(* IEC 61131-3 sources: 2026_Projet_YGO_ExcavatriceDragage/CODE/M_MAIN (part 2) *)

M1WinchSensors.CablePosM          := PRG_02_Acquisition.Data.EncoderM1.Measurement.CablePosM;
M1WinchSensors.Homed              := PRG_02_Acquisition.Data.EncoderM1.Homed;
M1WinchSensors.HomingSuspect      := PRG_02_Acquisition.Data.EncoderM1.HomingSuspect;
M1WinchSensors.ContactorsAllOff   := PRG_02_Acquisition.HwIn.Winch.M1_ContactorsReleased_DI;
M1WinchSensors.MeasuredSpeedBand  := instWinchLoadEstimatorM1.SpeedBand;
// Garde-fou vitesse mesuree : DESACTIVE par defaut (AF_Partie-10 §9bis, FB_Winch_v2.1 /
// FB_SpeedStep_v1.0 SpeedGuardEnable := FALSE). Le TRUE code en dur etait un reste de
// mise en service : il rendait la capacite de palier otage de instWinchSync (tout ecart
// sync -> SpeedGuardReady=FALSE -> clamp palier 1, y compris en montee).
// ⚠️ DETTE SAFETY -S5 : le garde-fou vitesse mesuree est HORS SERVICE. Le FB de
// gouvernance nominale annonce (FB_WinchRateInterlock) n'existe PAS dans CODE/.
// Decision : risque ACTE et documente — la surveillance survitesse reelle est portee par
// FB_Safety_Winch (gelee : harnais VAR_IN_OUT indisponible). Ne PAS armer une
// survitesse sur une table non prouvee. A re-trancher a la livraison .
// ⚠️ tache est BLOQUE (contrat C4 TASK_CONTRACT_AUTORITE_2_INTERLOCKS.yaml,
// ARRET VALIDATION HUMAINE requis : autorite, T_max/DropConfirmDelay, classification
// Fault.Error, argument PLr ; prerequis// non livres). Ne PAS creer
// FB_WinchRateInterlock hors de ce contrat — la logique de garde-fou existe deja dans
// FB_Winch §5 et reste volontairement desactivee (SpeedGuardEnable := FALSE) tant que la
// table SpeedBandMaxMps n'est pas validee en charge reelle (AF-10 §7.3 TBD).
M1WinchSensors.SpeedGuardEnable   := FALSE;
M1WinchSensors.SpeedGuardReady    := NOT instWinchSync.Fault.Error;

M1WinchCfg.SpeedStepTable         := _WinchSpeedStepTable;
M1WinchCfg.SlowdownDistanceTop_M  := _CommunCfgPersist.WinchSlowdownDistanceTop_M;
M1WinchCfg.SlowdownDistanceBottom_M := _CommunCfgPersist.WinchSlowdownDistanceBottom_M;
M1WinchCfg.SlowdownMaxStep        := _CommunCfgPersist.WinchSlowdownMaxStep;
// Cadence/interlocks : descente normale 500 ms, inversion vers descente 500 ms,
// montee normale 700 ms, inversion vers montee 800 ms.
// Champs non portes par la persistante -> assignes explicitement (le defaut de type n'est
// pas applique au runtime pour ce VAR local de struct). 0,7 s montee / 0,5 s descente.
M1WinchCfg.DirectionInterlockDelayAscent  := T#800ms;
M1WinchCfg.DirectionInterlockDelayDescent := T#500ms;
M1WinchCfg.StepRampDelayAscent    := T#700ms;
M1WinchCfg.StepRampDelayDescent   := T#500ms;

instWinchM1(
    Enable                  := (PRG_03_Modes_Cycle.Data.Auth.Mode <> E_Mode.DISABLE) AND NOT PRG_03_Modes_Cycle.Data.Auth.InhibitM1,
    Reset                   := PRG_07_Supervision.FaultMachineReset_IHM,
    PowerContactorEngaged   := PRG_02_Acquisition.HwIn.Machine.PowerContactorEngaged_DI,
    SafeStop                := SafeStopM1_Active,
    DescendPermit           := EffectivePermitM1_Descend,
    AscentPermit            := EffectivePermitM1_Ascent,
    WinchRequest            := ReqM1Winch,
    Sensors                 := M1WinchSensors,
    Config                  := M1WinchCfg,
    // ContactorFeedback (n°3 de la matrice) et Global — sans gate de mode (dérogation MES 2026).
    BypassContactorCheck    := (GVL_IHM.M1TreuilRetenue.Bypass.Global OR GVL_IHM.M1TreuilRetenue.Bypass.ContactorFeedback),
    BypassGlobal            := GVL_IHM.M1TreuilRetenue.Bypass.Global
);

// --- M2 : assemblage des structs ---
ReqM2Winch.RunRequest               := M2LogicRunRequest;
ReqM2Winch.ReqAscent                := M2LogicReqAscent;
ReqM2Winch.ReqDescend               := M2LogicReqDescend;
ReqM2Winch.SpeedStepReq             := M2LogicRequestStepTgt;
// Clamp de palier agrégé en §5ter : bornes communes M1=M2 (CommonMaxStep*) puis
// M2-propre (M2MaxStep*) — M2_BucketJogLimit / ManualBucketLimitsActive ne réduisent
// jamais M1 (pilotage unitaire M2). BucketNotClosedAscentCapStep1 /
// SlackCableAscentCapStep1 : réduisent M1 aussi UNIQUEMENT en pilotage couplé
// (CoupledBoth) — les 2 treuils liés doivent rester au même palier.
// D13 : reconstruction de table M2 supprimée — le clamp M2MaxStep* := 1 suffit
// (StepNumber ≤ 1 → seuls les états P1 sont commandés).
ReqM2Winch.MaxStepUp                := M2MaxStepUp;
ReqM2Winch.MaxStepDown              := M2MaxStepDown;
// Plancher palier descente plongée Kobold : plancher M2-propre agrégé en §5ter, injecté
// sur la cible (jamais sur StepNumber). Aucun effet si StartStop=FALSE.
ReqM2Winch.MinStepDown              := M2MinStepDown;
ReqM2Winch.HomingApproachActive     := PRG_03_Modes_Cycle.Data.Auth.HomingApproachEnable;
// Même limite haute active que FB_Safety_Winch (M2_LimitShift conservé).
ReqM2Winch.TopLimitM                := TopLimitM2_M;
ReqM2Winch.BottomLimitM             := BottomLimitM2_Active;
ReqM2Winch.SyncCoupled              := instWinchSync.SyncActive;

// === ATOMICITE DU DEMARRAGE COUPLE (volet M2, symetrique du volet M1 ~ligne 1225) ===
// Meme verrou : en intention both, si l'un des deux treuils n'est pas pret, on fige AUSSI
// la commande finale M2. Cas symetrique du REX : M2 relance seul pendant que M1 est en
// dead-time D18 -> cable qui file. On fige M2 UNIQUEMENT si M1 est le treuil pas pret.
IF NOT MaintN2 AND WinchBothMotionActive AND (instWinchM1.DirectionChangePending OR instWinchM1.Fault.Latched) THEN
    ReqM2Winch.RunRequest := FALSE; ReqM2Winch.ReqAscent := FALSE; ReqM2Winch.ReqDescend := FALSE; ReqM2Winch.SpeedStepReq := 0;
END_IF;

M2WinchSensors.CablePosM          := PRG_02_Acquisition.Data.EncoderM2.Measurement.CablePosM;
M2WinchSensors.Homed              := PRG_02_Acquisition.Data.EncoderM2.Homed;
M2WinchSensors.HomingSuspect      := PRG_02_Acquisition.Data.EncoderM2.HomingSuspect;
M2WinchSensors.ContactorsAllOff   := PRG_02_Acquisition.HwIn.Winch.M2_ContactorsReleased_DI;
M2WinchSensors.MeasuredSpeedBand  := instWinchLoadEstimatorM2.SpeedBand;
// Garde-fou vitesse mesuree : DESACTIVE par defaut (idem M1 ci-dessus, AF_Partie-10 §9bis).
M2WinchSensors.SpeedGuardEnable   := FALSE;
M2WinchSensors.SpeedGuardReady    := NOT instWinchSync.Fault.Error;

M2WinchCfg.SpeedStepTable         := _WinchSpeedStepTable;
M2WinchCfg.SlowdownDistanceTop_M  := _CommunCfgPersist.WinchSlowdownDistanceTop_M;
M2WinchCfg.SlowdownDistanceBottom_M := _CommunCfgPersist.WinchSlowdownDistanceBottom_M;
M2WinchCfg.SlowdownMaxStep        := _CommunCfgPersist.WinchSlowdownMaxStep;
// Cadence/interlocks identiques M1 : descente normale 500 ms, inversion vers descente
// 500 ms, montee normale 700 ms, inversion vers montee 800 ms.
M2WinchCfg.DirectionInterlockDelayAscent  := T#800ms;
M2WinchCfg.DirectionInterlockDelayDescent := T#500ms;
M2WinchCfg.StepRampDelayAscent    := T#700ms;
M2WinchCfg.StepRampDelayDescent   := T#500ms;

instWinchM2(
    Enable                  := (PRG_03_Modes_Cycle.Data.Auth.Mode <> E_Mode.DISABLE) AND NOT PRG_03_Modes_Cycle.Data.Auth.InhibitM2,
    Reset                   := PRG_07_Supervision.FaultMachineReset_IHM,
    PowerContactorEngaged   := PRG_02_Acquisition.HwIn.Machine.PowerContactorEngaged_DI,
    SafeStop                := SafeStopM2_Active,
    DescendPermit           := M2DescendPermitApplied,
    AscentPermit            := M2AscentPermitApplied,
    WinchRequest            := ReqM2Winch,
    Sensors                 := M2WinchSensors,
    Config                  := M2WinchCfg,
    // Idem M1 ci-dessus
    BypassContactorCheck    := (GVL_IHM.M2TreuilBenne.Bypass.Global OR GVL_IHM.M2TreuilBenne.Bypass.ContactorFeedback),
    BypassGlobal            := GVL_IHM.M2TreuilBenne.Bypass.Global
);

// Atomicite de sortie couplee : les deux FB_Winch ont maintenant traite la demande du
// scan. Leur readiness directionnelle courante est donc connue avant publication vers
// PRG_06. La barriere finale ne recevra aucun relais/contacteur tant qu'un axe attend.
WinchBothMotionReady := NOT (instWinchM1.DirectionChangePending OR instWinchM2.DirectionChangePending)
                        AND NOT instWinchM1.Fault.Latched AND NOT instWinchM2.Fault.Latched;

// ── Collecteurs passifs d'apprentissage vitesse par palier ──
// Appelés APRÈS instWinchM1/M2 : StepNumber lu = palier courant du scan (pas de lag).
// Dérivations des entrées de collecte :
//   • LoadPresent : charge présente si l'estimateur de charge (même source vitesse) estime
//     une charge >= 50 % (seuil de mise en service, à confirmer sur site).
//   • StableForLearn : treuil commandé (palier > 0) et sans défaut — conditions stables.
// Collecteur STRICTEMENT PASSIF : aucune commande moteur, aucune surveillance survitesse
// (la survitesse reste, gelée — voir bandeau §6 M1/M2 SpeedGuardEnable).
LoadPresentM1 := (instWinchLoadEstimatorM1.EstimatedLoadPct >= 50.0);
LoadPresentM2 := (instWinchLoadEstimatorM2.EstimatedLoadPct >= 50.0);
StableForLearnM1 := (instWinchM1.StepNumber > 0) AND NOT instWinchM1.Fault.Error;
StableForLearnM2 := (instWinchM2.StepNumber > 0) AND NOT instWinchM2.Fault.Error;

instWinchSpeedLearningM1(
    Enable              := (PRG_03_Modes_Cycle.Data.Auth.Mode <> E_Mode.DISABLE) AND NOT PRG_03_Modes_Cycle.Data.Auth.InhibitM1,
    LearnStart          := GVL_IHM.M1TreuilRetenue.Cmd.BtnLearnSpeed,
    WinchId             := 1,
    ReqAscent          := M1LogicReqAscent,
    ReqDescend         := M1LogicReqDescend,
    StepNumber          := instWinchM1.StepNumber,
    MeasuredSpeedMps    := PRG_02_Acquisition.Data.EncoderM1.Measurement.Speed_Mps,
    MeasuredSpeedValid  := PRG_02_Acquisition.Data.EncoderM1.Measurement.SpeedValid,
    LoadPresent         := LoadPresentM1,
    StableForLearn      := StableForLearnM1,
    Config              := _WinchSpeedLearnCfg,
    Table               := _WinchSpeedLearnTable
);

instWinchSpeedLearningM2(
    Enable              := (PRG_03_Modes_Cycle.Data.Auth.Mode <> E_Mode.DISABLE) AND NOT PRG_03_Modes_Cycle.Data.Auth.InhibitM2,
    LearnStart          := GVL_IHM.M2TreuilBenne.Cmd.BtnLearnSpeed,
    WinchId             := 2,
    ReqAscent          := M2LogicReqAscent,
    ReqDescend         := M2LogicReqDescend,
    StepNumber          := instWinchM2.StepNumber,
    MeasuredSpeedMps    := PRG_02_Acquisition.Data.EncoderM2.Measurement.Speed_Mps,
    MeasuredSpeedValid  := PRG_02_Acquisition.Data.EncoderM2.Measurement.SpeedValid,
    LoadPresent         := LoadPresentM2,
    StableForLearn      := StableForLearnM2,
    Config              := _WinchSpeedLearnCfg,
    Table               := _WinchSpeedLearnTable
);

{endregion}

{region "📤 §7 Publication demandes"}
// === 📤 §7 PUBLICATION DEMANDES BRUTES (WinchM1/M2FinalInterlockRequest) ===

WinchM1FinalInterlockRequest.Enable := TRUE;
WinchM1FinalInterlockRequest.Reset := PRG_07_Supervision.FaultMachineReset_IHM;
WinchM1FinalInterlockRequest.PowerContactorEngaged := PRG_02_Acquisition.HwIn.Machine.PowerContactorEngaged_DI;
WinchM1FinalInterlockRequest.SafeStop := SafeStopM1_Active;
// Plus de BrakeReleaseRequest/
// BrakeCommandOpenConfirmed calcules par FB_Winch — la barriere finale
// (FB_WinchOutputInterlock) recoit le retour PHYSIQUE brut directement,
// et calcule elle-meme BrakeCmd := RelayFwd OR RelayRev (voir bandeau de ce FB).
WinchM1FinalInterlockRequest.BrakeFeedback := SEL(MaintN2 OR GVL_IHM.M1TreuilRetenue.Bypass.ContactorFeedback OR GVL_IHM.M1TreuilRetenue.Bypass.Global,
                                                   PRG_02_Acquisition.HwIn.Winch.M1_BrakeIsOpen_DI,
                                                   instWinchM1.RelayFwd OR instWinchM1.RelayRev);
WinchM1FinalInterlockRequest.FwdRevSpeedFeedbackOff := SEL(MaintN2 OR GVL_IHM.M1TreuilRetenue.Bypass.ContactorFeedback OR GVL_IHM.M1TreuilRetenue.Bypass.Global,
                                                           PRG_02_Acquisition.HwIn.Winch.M1_ContactorsReleased_DI,
                                                           NOT (instWinchM1.RelayFwd OR instWinchM1.RelayRev));
WinchM1FinalInterlockRequest.RequestedRelayFwd := instWinchM1.RelayFwd;
WinchM1FinalInterlockRequest.RequestedRelayRev := instWinchM1.RelayRev;
WinchM1FinalInterlockRequest.RequestedContactor1 := instWinchM1.Contactor1;
WinchM1FinalInterlockRequest.RequestedContactor2 := instWinchM1.Contactor2;
WinchM1FinalInterlockRequest.RequestedContactor3 := instWinchM1.Contactor3;
WinchM1FinalInterlockRequest.RequestedContactor4 := instWinchM1.Contactor4;
WinchM1FinalInterlockRequest.RequestedStep := instWinchM1.StepNumber;
WinchM1FinalInterlockRequest.PowerCutOff := instSafetyWinchM1.PowerCutOff;
WinchM1FinalInterlockRequest.AscentPermit := EffectivePermitM1_Ascent;
WinchM1FinalInterlockRequest.DescendPermit := EffectivePermitM1_Descend;

WinchM2FinalInterlockRequest.Enable := TRUE;
WinchM2FinalInterlockRequest.Reset := PRG_07_Supervision.FaultMachineReset_IHM;
WinchM2FinalInterlockRequest.PowerContactorEngaged := PRG_02_Acquisition.HwIn.Machine.PowerContactorEngaged_DI;
WinchM2FinalInterlockRequest.SafeStop := SafeStopM2_Active;
WinchM2FinalInterlockRequest.BrakeFeedback := SEL(MaintN2 OR GVL_IHM.M2TreuilBenne.Bypass.ContactorFeedback OR GVL_IHM.M2TreuilBenne.Bypass.Global,
                                                   PRG_02_Acquisition.HwIn.Winch.M2_BrakeIsOpen_DI,
                                                   instWinchM2.RelayFwd OR instWinchM2.RelayRev);
WinchM2FinalInterlockRequest.FwdRevSpeedFeedbackOff := SEL(MaintN2 OR GVL_IHM.M2TreuilBenne.Bypass.ContactorFeedback OR GVL_IHM.M2TreuilBenne.Bypass.Global,
                                                           PRG_02_Acquisition.HwIn.Winch.M2_ContactorsReleased_DI,
                                                           NOT (instWinchM2.RelayFwd OR instWinchM2.RelayRev));
WinchM2FinalInterlockRequest.RequestedRelayFwd := instWinchM2.RelayFwd;
WinchM2FinalInterlockRequest.RequestedRelayRev := instWinchM2.RelayRev;
WinchM2FinalInterlockRequest.RequestedContactor1 := instWinchM2.Contactor1;
WinchM2FinalInterlockRequest.RequestedContactor2 := instWinchM2.Contactor2;
WinchM2FinalInterlockRequest.RequestedContactor3 := instWinchM2.Contactor3;
WinchM2FinalInterlockRequest.RequestedContactor4 := instWinchM2.Contactor4;
WinchM2FinalInterlockRequest.RequestedStep := instWinchM2.StepNumber;
WinchM2FinalInterlockRequest.PowerCutOff := instSafetyWinchM2.PowerCutOff;
WinchM2FinalInterlockRequest.AscentPermit := M2AscentPermitApplied;
WinchM2FinalInterlockRequest.DescendPermit := M2DescendPermitApplied;

WinchBothFinalStep45Coherent :=
    PRG_03_Modes_Cycle.Data.AutoDiveM1Step4M2Step5Active
    AND NOT WinchM1FinalInterlockRequest.RequestedRelayFwd
    AND NOT WinchM2FinalInterlockRequest.RequestedRelayFwd
    AND WinchM1FinalInterlockRequest.RequestedRelayRev
    AND WinchM2FinalInterlockRequest.RequestedRelayRev
    AND (WinchM1FinalInterlockRequest.RequestedStep = 4)
    AND (WinchM2FinalInterlockRequest.RequestedStep = 5)
    AND (WinchM1FinalInterlockRequest.RequestedContactor1 = _WinchSpeedStepTable.P4R1)
    AND (WinchM1FinalInterlockRequest.RequestedContactor2 = _WinchSpeedStepTable.P4R2)
    AND (WinchM1FinalInterlockRequest.RequestedContactor3 = _WinchSpeedStepTable.P4R3)
    AND (WinchM1FinalInterlockRequest.RequestedContactor4 = _WinchSpeedStepTable.P4R4)
    AND (WinchM2FinalInterlockRequest.RequestedContactor1 = _WinchSpeedStepTable.P5R1)
    AND (WinchM2FinalInterlockRequest.RequestedContactor2 = _WinchSpeedStepTable.P5R2)
    AND (WinchM2FinalInterlockRequest.RequestedContactor3 = _WinchSpeedStepTable.P5R3)
    AND (WinchM2FinalInterlockRequest.RequestedContactor4 = _WinchSpeedStepTable.P5R4);

WinchBothFinalRequestsCoherent :=
    WinchBothFinalStep45Coherent
    OR ((WinchM1FinalInterlockRequest.RequestedRelayFwd = WinchM2FinalInterlockRequest.RequestedRelayFwd)
        AND (WinchM1FinalInterlockRequest.RequestedRelayRev = WinchM2FinalInterlockRequest.RequestedRelayRev)
        AND (WinchM1FinalInterlockRequest.RequestedContactor1 = WinchM2FinalInterlockRequest.RequestedContactor1)
        AND (WinchM1FinalInterlockRequest.RequestedContactor2 = WinchM2FinalInterlockRequest.RequestedContactor2)
        AND (WinchM1FinalInterlockRequest.RequestedContactor3 = WinchM2FinalInterlockRequest.RequestedContactor3)
        AND (WinchM1FinalInterlockRequest.RequestedContactor4 = WinchM2FinalInterlockRequest.RequestedContactor4)
        AND (WinchM1FinalInterlockRequest.RequestedStep = WinchM2FinalInterlockRequest.RequestedStep));

// Defense en profondeur apres les deux FB : en intention couplee, aucun actionneur ne
// peut etre publie seul. Les FB continuent d'evaluer leurs interlocks internes, mais les
// deux demandes physiques restent neutres jusqu'a readiness commune.
IF (PRG_03_Modes_Cycle.Data.Auth.Mode = E_Mode.SEMI_AUTO)
   AND WinchBothMotionActive
   AND (NOT WinchBothMotionReady OR NOT WinchBothFinalRequestsCoherent) THEN
    WinchM1FinalInterlockRequest.RequestedRelayFwd := FALSE;
    WinchM1FinalInterlockRequest.RequestedRelayRev := FALSE;
    WinchM1FinalInterlockRequest.RequestedContactor1 := FALSE;
    WinchM1FinalInterlockRequest.RequestedContactor2 := FALSE;
    WinchM1FinalInterlockRequest.RequestedContactor3 := FALSE;
    WinchM1FinalInterlockRequest.RequestedContactor4 := FALSE;
    WinchM1FinalInterlockRequest.RequestedStep := 0;
    WinchM2FinalInterlockRequest.RequestedRelayFwd := FALSE;
    WinchM2FinalInterlockRequest.RequestedRelayRev := FALSE;
    WinchM2FinalInterlockRequest.RequestedContactor1 := FALSE;
    WinchM2FinalInterlockRequest.RequestedContactor2 := FALSE;
    WinchM2FinalInterlockRequest.RequestedContactor3 := FALSE;
    WinchM2FinalInterlockRequest.RequestedContactor4 := FALSE;
    WinchM2FinalInterlockRequest.RequestedStep := 0;
END_IF;

{endregion}

{region "📊 §8 Publication états IHM"}
// === 📤 §8 PUBLICATION ÉTATS IHM (faits publics, lecture seule) ===
// Projection déléguée à FB_WinchStateProjection () : recopie bit-identique
// des sources → WinchM1State/WinchM2State/WinchM1Safety/WinchM2Safety/CableLimitAscent.
// Aucune logique de commande modifiée (non-régression). SyncState/BucketState/
// Benne_IsRoughlyClosed/GLV_IHM restent ici (hors scope du FB).
instWinchStateProjection(
    EncoderM1 := PRG_02_Acquisition.Data.EncoderM1,
    EncoderM2 := PRG_02_Acquisition.Data.EncoderM2,
    WinchM1Ref := instWinchM1,
    WinchM2Ref := instWinchM2,
    SafetyM1 := instSafetyWinchM1,
    SafetyM2 := instSafetyWinchM2,
    InterlockM1 := PRG_06_Outputs.instWinchOutputInterlockM1,
    InterlockM2 := PRG_06_Outputs.instWinchOutputInterlockM2,
    Auth := PRG_03_Modes_Cycle.Data.Auth,
    HwInWinch := PRG_02_Acquisition.HwIn.Winch,
    HwRealWinch := PRG_02_Acquisition.HwReal.Winch,
    M1_PrevSpeed_Mps := M1_PrevSpeed_Mps,
    M2_PrevSpeed_Mps := M2_PrevSpeed_Mps,
    M1LogicRequestSpeedCmd_Pct := M1LogicRequestSpeedCmd_Pct,
    M2LogicRequestSpeedCmd_Pct := M2LogicRequestSpeedCmd_Pct,
    BottomLimitM1_Active := BottomLimitM1_Active,
    BottomLimitM2_Active := BottomLimitM2_Active,
    SafeStopM1_Active := SafeStopM1_Active,
    SafeStopM2_Active := SafeStopM2_Active,
    EffectivePermitM1_Ascent := EffectivePermitM1_Ascent,
    EffectivePermitM1_Descend := EffectivePermitM1_Descend,
    EffectivePermitM2_Ascent := EffectivePermitM2_Ascent,
    EffectivePermitM2_Descend := EffectivePermitM2_Descend,
    M2_LimitShift := M2_LimitShift,
    CfgCableLimitAscent_M := _CommunCfgPersist.CfgCableLimitAscent_M,
    CfgCableLimitDescentM1_M := _WinchM1CfgPersist.CfgCableLimitDescent_M,
    CfgCableLimitDescentM2_M := _WinchM2CfgPersist.CfgCableLimitDescent_M,
    EncoderM1_Operational := PRG_02_Acquisition.Data.Network.EncoderM1.Operational,
    EncoderM2_Operational := PRG_02_Acquisition.Data.Network.EncoderM2.Operational,
    M1PowerCutOffSafetyInfo := PRG_06_Outputs.M1PowerCutOffSafetyInfo,
    M1SafeStopSafetyInfo := PRG_06_Outputs.M1SafeStopSafetyInfo,
    M1BlockedBySafetyInfo := PRG_06_Outputs.M1BlockedBySafetyInfo,
    M2PowerCutOffSafetyInfo := PRG_06_Outputs.M2PowerCutOffSafetyInfo,
    M2SafeStopSafetyInfo := PRG_06_Outputs.M2SafeStopSafetyInfo,
    M2BlockedBySafetyInfo := PRG_06_Outputs.M2BlockedBySafetyInfo
);
WinchM1State := instWinchStateProjection.WinchM1State;
WinchM2State := instWinchStateProjection.WinchM2State;
WinchM1Safety := instWinchStateProjection.WinchM1Safety;
WinchM2Safety := instWinchStateProjection.WinchM2Safety;
CableLimitAscentM1Reached := instWinchStateProjection.CableLimitAscentM1Reached;
CableLimitAscentM2Reached := instWinchStateProjection.CableLimitAscentM2Reached;

SyncState.DeltaPos_M := instWinchSync.SignedDeltaPosM;
SyncState.SyncActive := instWinchSync.SyncActive;
SyncState.SyncWarn := instWinchSync.SyncWarn;
SyncState.SyncDeviationWarn := instWinchSync.SyncDeviationWarn;
SyncState.Ready := instWinchSync.Ready;
SyncState.Error := instWinchSync.Fault.Error;
SyncState.FaultLatched := instWinchSync.Fault.Latched;
SyncState.ErrorId := instWinchSync.Fault.ErrorId;
IF instWinchSync.Fault.Error THEN
    SyncState.FBState := E_State.ERROR;
ELSIF instWinchSync.SyncActive THEN
    SyncState.FBState := E_State.BUSY;
ELSE
    SyncState.FBState := E_State.READY;
END_IF;

BucketState.MechState := _BucketState;
BucketState.MechState.ActiveOffsetValid := instBucket.ActiveOffsetValid;
IF instBucket.Fault.Error THEN
    BucketState.FBState := E_State.ERROR;
ELSIF instBucket.Lifecycle.Busy THEN
    BucketState.FBState := E_State.BUSY;
ELSE
    BucketState.FBState := E_State.READY;
END_IF;
BucketState.ActiveOffset_M := instBucket.ActiveOffsetM;
BucketState.M2RunRequest := instBucket.M2_RunRequest;
BucketState.M2ReqAscent := instBucket.M2_ReqAscent;
BucketState.M2ReqDescend := instBucket.M2_ReqDescend;
BucketState.M2BucketJogLimit := instBucket.M2_BucketJogLimit;
BucketState.ManualBucketLimitsActive := ManualBucketLimitsActive;
BucketState.OffsetStateMismatchWarn := instBucket.OffsetStateMismatchWarn;
// Affichage operateur (bargraphe) et traces (T291-B) : DisplayOffsetM continu
// (LIMIT OffsetOpenM..OffsetCloseM), pas de saut de 15 m aux transitions d'états francs.
BucketState.M2PositionCorrected := PRG_02_Acquisition.Data.EncoderM2.Measurement.CablePosM - instBucket.DisplayOffsetM;
// Qualification mesure indépendante : conservateur (T291-B B1). En position intermédiaire,
// la mesure absorbe la dérive propre de M2 -> M2PositionCorrectedValid reste FALSE pour
// interdire tout usage FDC/safety. Seuls les états francs stabilisés (IsClosed XOR IsOpen)
// avec benne référencée sont qualifiés pour la surveillance indépendante.
BucketState.M2PositionCorrectedValid := _BucketState.BucketReferenced
    AND (_BucketState.IsClosed XOR _BucketState.IsOpen);
BucketState.Ready := instBucket.Ready;
BucketState.Busy := instBucket.Lifecycle.Busy;
BucketState.Done := instBucket.Lifecycle.Done;
Data.BucketCloseReached := instBucket.CloseReached;
BucketState.Error := instBucket.Fault.Error;
BucketState.FaultLatched := instBucket.Fault.Latched;
BucketState.ErrorId := instBucket.Fault.ErrorId;
BucketState.RemainingTravel_M := instBucket.RemainingTravelM;
BucketState.DeltaPosition_M := instBucket.DeltaPosition_M;
BucketState.DeltaPositionCorrected_M := instBucket.DeltaPositionCorrected_M;
BucketState.BucketOpening_Pct := instBucket.BucketOpening_Pct;
BucketState.CloseActive := instBucket.CloseReq;
BucketState.OpenActive := instBucket.OpenReq;
// Reflète le séquencement auto : occupé sur une ouverture/fermeture qu'IL a armée, ou en phase
// vitesse contrôlée post-fermeture.
BucketState.AutoBucketSeqActive := (instBucket.Lifecycle.Busy AND (WinchBothDiveBucketOpenArmed OR WinchBothAscentBucketCloseArmed)) OR ExtractionControlActive;
BucketState.CoupledDiveOpenArmed := WinchBothDiveBucketOpenArmed;
BucketState.CoupledAscentCloseArmed := WinchBothAscentBucketCloseArmed;
BucketState.MachineHomed := PRG_02_Acquisition.Data.MachineHoming.Homed;
BucketState.MachineHomingStep := PRG_02_Acquisition.Data.MachineHoming.Step;
BucketState.MachineHomingInstruction := PRG_02_Acquisition.Data.MachineHoming.Instruction;
BucketState.MachineHomingFailed := PRG_02_Acquisition.Data.MachineHoming.Failed;
BucketState.MachineHomingActive := PRG_02_Acquisition.Data.MachineHoming.Active;
BucketState.MachineHomingLossSafeStop := PRG_02_Acquisition.Data.MachineHoming.HomingLoss;
BucketState.ExtractionControlActive := ExtractionControlActive;
BucketState.CoupledMotionBlockedByBucket := WinchBothMotionBlockedByBucket;
GVL_IHM.Commun.KoboldImmersionConfirmed := KoboldImmersionConfirmed;
GVL_IHM.Commun.KoboldBottomTouchLatched := KoboldBottomTouchLatched;

// Tolérance matière benne : « à peu près fermée » = fermée OU
// intermédiaire proche de l'offset fermé (tolérance 2 m). Évite le blocage au fond sur
// matière dense (galets) qui ne ferme jamais à 100% de la consigne fine.
// 🎛️ Branche AJOUTÉE, jamais substitutive : la ligne 2 m ci-dessous est INTOUCHÉE (valeur,
// sens et rôle de filet anti-blocage conservés). La disjonction ajoutée permet d'avancer
// l'instant où la fermeture est considérée atteinte, via le réglage d'ouverture benne
// (0 = branche inactive -> critère d'arrivée seul).
// Mesure QUALIFIÉE identique à celle de FB_Bucket (références M1/M2, absence de défaut
// latché — géométrie benne invalide incluse — et référence benne persistante) : le même
// signal des deux côtés, sinon la fenêtre de sortie AX10 pourrait se refermer entre les
// deux évaluations et figer la séquence.
ThresholdMeasureValid := PRG_02_Acquisition.Data.EncoderM1.Homed
                         AND PRG_02_Acquisition.Data.EncoderM2.Homed
                         AND NOT instBucket.Fault.Error
                         AND _BucketState.BucketReferenced;
instCloseThreshold(
    ThresholdPct    := GVL_IHM.CycleSemiAuto.Cfg.ExtractionStartOpening_Pct,
    OffsetOpenM     := _BucketCfgPersist.Config.OffsetOpenM,
    OffsetCloseM    := _BucketCfgPersist.Config.OffsetCloseM,
    DeltaPosition_M := instBucket.DeltaPosition_M,
    MeasureValid    := ThresholdMeasureValid,
    IsIntermediate  := _BucketState.IsIntermediate
);
Benne_IsRoughlyClosed := _BucketState.IsClosed
    OR (_BucketState.IsIntermediate
        AND (instBucket.DeltaPosition_M >= (_BucketCfgPersist.Config.OffsetCloseM - 2.0)))
    OR instCloseThreshold.Reached;

{region "🕵️ §8bis Trace blocage"}
// === 🕵️ §8bis TRACE DE BLOCAGE TERRAIN (cause priorisée + horodatage) ===
// Diagnostic lecture seule, publié via Data.TraceM1/M2 et consommé par FB_TroubleshootingView.
// L'ordre IF/ELSIF EST l'ordre de priorité (cf. E_WinchTraceBlockReason) : la cause la plus
// grave gagne. BlockReasonTimestamp est latched au premier scan du changement (1 scan, mémoire).
// Aucune action de conduite ne dépend de ces champs.

// --- M1 ---
TraceM1.DescendPermitEffective := EffectivePermitM1_Descend;
TraceM1.AscentPermitEffective  := EffectivePermitM1_Ascent;
TraceM1.AscentPermitApplied     := EffectivePermitM1_Ascent;
TraceM1.DescendPermitApplied    := EffectivePermitM1_Descend;
TraceM1.FinalPermitBlocked      := (ReqM1Winch.RunRequest AND ReqM1Winch.ReqAscent AND NOT EffectivePermitM1_Ascent)
                               OR (ReqM1Winch.RunRequest AND ReqM1Winch.ReqDescend AND NOT EffectivePermitM1_Descend);
TraceM1.SafeStopActive         := SafeStopM1_Active;
TraceM1.SafeStopSourceSafety   := instSafetyWinchM1.SafeStop;
TraceM1.SafeStopSourceInput    := PRG_02_Acquisition.Data.InputModules.Fault
                                  OR PRG_02_Acquisition.Data.MachineHoming.HomingLoss
                                  OR instBucket.M1SlipDetected;
TraceM1.SafeStopSourceSync     := ((instWinchSync.Fault.ErrorId AND 16#0002) <> 16#0000)
                                  OR (instWinchSync.SyncActive AND SafeStopM2_Raw);
TraceM1.PowerCutOffActive      := instSafetyWinchM1.PowerCutOff;
TraceM1.Inhibited              := (PRG_03_Modes_Cycle.Data.Auth.Mode = E_Mode.DISABLE)
                                  OR PRG_03_Modes_Cycle.Data.Auth.InhibitM1;
TraceM1.FinalInterlockError    := WinchM1State.FinalInterlockError;
TraceM1.FinalInterlockReason   := WinchM1State.FinalInterlockReason;
TraceM1.StepNumber             := WinchM1State.StepNumber;

IF instSafetyWinchM1.PowerCutOff THEN
    TraceM1.BlockReason := E_WinchTraceBlockReason.POWER_CUTOFF;
ELSIF TraceM1.Inhibited THEN
    TraceM1.BlockReason := E_WinchTraceBlockReason.AXIS_DISABLED;
ELSIF SafeStopM1_Active THEN
    TraceM1.BlockReason := E_WinchTraceBlockReason.SAFESTOP;
ELSIF instSafetyWinchM1.Fault.Error THEN
    TraceM1.BlockReason := E_WinchTraceBlockReason.SAFETY_FAULT;
ELSIF NOT (SafetyPermitM1_Ascent OR SafetyPermitM1_Descend) THEN
    TraceM1.BlockReason := E_WinchTraceBlockReason.SAFETY_PERMIT_MISSING;
ELSIF NOT (ProcessPermitM1_Ascent OR ProcessPermitM1_Descend) THEN
    TraceM1.BlockReason := E_WinchTraceBlockReason.PROCESS_PERMIT_MISSING;
ELSIF NOT (EffectivePermitM1_Ascent OR EffectivePermitM1_Descend) THEN
    TraceM1.BlockReason := E_WinchTraceBlockReason.COUPLING_BLOCKED;
ELSIF instWinchM1.Fault.Error THEN
    TraceM1.BlockReason := E_WinchTraceBlockReason.WINCH_FAULT;
ELSIF WinchM1State.FinalInterlockError THEN
    TraceM1.BlockReason := E_WinchTraceBlockReason.FINAL_INTERLOCK_BLOCKED;
ELSE
    TraceM1.BlockReason := E_WinchTraceBlockReason.NONE;
END_IF;
IF TraceM1.BlockReason <> TraceM1_PrevReason THEN
    TraceM1.BlockReasonTimestamp := TIME_TO_UDINT(TIME());
END_IF;
TraceM1_PrevReason := TraceM1.BlockReason;

// --- M2 ---
TraceM2.DescendPermitEffective := EffectivePermitM2_Descend;
TraceM2.AscentPermitEffective  := EffectivePermitM2_Ascent;
TraceM2.AscentPermitApplied     := M2AscentPermitApplied;
TraceM2.DescendPermitApplied    := M2DescendPermitApplied;
TraceM2.FinalPermitBlocked      := (ReqM2Winch.RunRequest AND ReqM2Winch.ReqAscent AND NOT EffectivePermitM2_Ascent)
                               OR (ReqM2Winch.RunRequest AND ReqM2Winch.ReqDescend AND NOT EffectivePermitM2_Descend);
TraceM2.SafeStopActive         := SafeStopM2_Active;
TraceM2.SafeStopSourceSafety   := instSafetyWinchM2.SafeStop;
TraceM2.SafeStopSourceInput    := PRG_02_Acquisition.Data.InputModules.Fault
                                  OR PRG_02_Acquisition.Data.MachineHoming.HomingLoss;
TraceM2.SafeStopSourceSync     := ((instWinchSync.Fault.ErrorId AND 16#0002) <> 16#0000)
                                  OR (instWinchSync.SyncActive AND SafeStopM1_Raw);
TraceM2.PowerCutOffActive      := instSafetyWinchM2.PowerCutOff;
TraceM2.Inhibited              := (PRG_03_Modes_Cycle.Data.Auth.Mode = E_Mode.DISABLE)
                                  OR PRG_03_Modes_Cycle.Data.Auth.InhibitM2;
TraceM2.FinalInterlockError    := WinchM2State.FinalInterlockError;
TraceM2.FinalInterlockReason   := WinchM2State.FinalInterlockReason;
TraceM2.StepNumber             := WinchM2State.StepNumber;

IF instSafetyWinchM2.PowerCutOff THEN
    TraceM2.BlockReason := E_WinchTraceBlockReason.POWER_CUTOFF;
ELSIF TraceM2.Inhibited THEN
    TraceM2.BlockReason := E_WinchTraceBlockReason.AXIS_DISABLED;
ELSIF SafeStopM2_Active THEN
    TraceM2.BlockReason := E_WinchTraceBlockReason.SAFESTOP;
ELSIF instSafetyWinchM2.Fault.Error THEN
    TraceM2.BlockReason := E_WinchTraceBlockReason.SAFETY_FAULT;
ELSIF NOT (SafetyPermitM2_Ascent OR SafetyPermitM2_Descend) THEN
    TraceM2.BlockReason := E_WinchTraceBlockReason.SAFETY_PERMIT_MISSING;
ELSIF NOT (ProcessPermitM2_Ascent OR ProcessPermitM2_Descend) THEN
    TraceM2.BlockReason := E_WinchTraceBlockReason.PROCESS_PERMIT_MISSING;
ELSIF NOT (EffectivePermitM2_Ascent OR EffectivePermitM2_Descend) THEN
    TraceM2.BlockReason := E_WinchTraceBlockReason.COUPLING_BLOCKED;
ELSIF instWinchM2.Fault.Error THEN
    TraceM2.BlockReason := E_WinchTraceBlockReason.WINCH_FAULT;
ELSIF WinchM2State.FinalInterlockError THEN
    TraceM2.BlockReason := E_WinchTraceBlockReason.FINAL_INTERLOCK_BLOCKED;
ELSE
    TraceM2.BlockReason := E_WinchTraceBlockReason.NONE;
END_IF;
IF TraceM2.BlockReason <> TraceM2_PrevReason THEN
    TraceM2.BlockReasonTimestamp := TIME_TO_UDINT(TIME());
END_IF;
TraceM2_PrevReason := TraceM2.BlockReason;

{endregion}

// 🧩 Cause de blocage priorisée sur l'état public IHM (miroir de la trace terrain §8bis)
WinchM1State.AxisBlockReason := TraceM1.BlockReason;
WinchM2State.AxisBlockReason := TraceM2.BlockReason;

// === 🔌 PUBLICATION BUS INTER-PRG (Data : ST_WinchInterPrg) ===
// Copie des structs internes vers le bus de sortie (producteur unique).
Data.WinchM1FinalInterlockRequest := WinchM1FinalInterlockRequest;
Data.WinchM2FinalInterlockRequest := WinchM2FinalInterlockRequest;
Data.M1LogicRequestSpeedCmd_Pct   := M1LogicRequestSpeedCmd_Pct;
Data.M2LogicRequestSpeedCmd_Pct   := M2LogicRequestSpeedCmd_Pct;
Data.KoboldContactorCmdArbitrated := KoboldContactorCmdArbitrated;
Data.WinchM1State                 := WinchM1State;
Data.WinchM2State                 := WinchM2State;
Data.WinchM1Safety                := WinchM1Safety;
Data.WinchM2Safety                := WinchM2Safety;
Data.SyncState                    := SyncState;
// Signal BLOQUANT unique du cycle : le bit 0 Fault.Error est un simple warning
// (degradation palier 1), il ne doit jamais faire basculer le grafcet en AX_STAB.
// Les protections critiques restent : deviation confirmee, contacteurs, et Meca E.
Data.WinchSyncError               := instWinchSync.SyncDeviationFault
                                     OR instWinchSync.ContactorMismatch
                                     OR WinchM1Safety.ErrorMecaE
                                     OR WinchM2Safety.ErrorMecaE;
Data.WinchSyncSignedDeltaPosM     := instWinchSync.SignedDeltaPosM;
Data.AutoDiveM1Step4M2Step5Active := PRG_03_Modes_Cycle.Data.AutoDiveM1Step4M2Step5Active;
Data.BucketState                  := BucketState;
Data.Benne_IsRoughlyClosed        := Benne_IsRoughlyClosed;
Data.BucketBusy                   := instBucket.Lifecycle.Busy;
Data.BucketDone                   := instBucket.Lifecycle.Done;
Data.BucketError                  := instBucket.Fault.Error;
Data.EffectivePermitBucket_Open   := EffectivePermitBucket_Open;
Data.EffectivePermitBucket_Close  := EffectivePermitBucket_Close;
Data.ArmingPermit                 := ArmingPermit;
Data.ProcessPermitM1_Ascent       := ProcessPermitM1_Ascent;
Data.ProcessPermitM1_Descend      := ProcessPermitM1_Descend;
Data.ProcessPermitM2_Ascent       := ProcessPermitM2_Ascent;
Data.ProcessPermitM2_Descend      := ProcessPermitM2_Descend;
Data.DescendPermitDiveBucketOpen  := DescendPermitDiveBucketOpen;
Data.ExtractionAssistActive       := ExtractionAssistActive;
Data.ExtractionAscentPermit       := PRG_03_Modes_Cycle.Data.ReqProgram.ReqBucket.AscentPermit;
// Usage effectif d'un override/bypass de position (consommé PRG_03 → FB_Modes)
Data.PositionLimitOverriddenM1    := PositionLimitOverriddenM1;
Data.PositionLimitOverriddenM2    := PositionLimitOverriddenM2;
// 🕵️ Trace de blocage terrain (consommée FB_TroubleshootingView)
Data.TraceM1                      := TraceM1;
Data.TraceM2                      := TraceM2;
// 🔗 ATOMICITÉ BOTH : diagnostic IHM lecture seule
Data.BothActive                   := WinchBothMotionActive;
Data.BothBlocked                  := BothBlocked;
Data.BothBlockReason              := BothBlockReason;

{endregion}
END_PROGRAM

(* ---- PRG_05_Translation.st ---- *)
(* ═══════════════════════════════════════════════════════════════
   ↔️ PRG_05_Translation — Pilotage de la Translation M3
   ───────────────────────────────────────────────────────────────
   ⚙️ Exécuté par la tâche PLC en position 5 (après PRG_04_Treuils_Benne).
   ✅ Arbitre entre les commandes Manuelles (Joystick) et Automatiques (PRG_03_Modes_Cycle).
   📄 Docs : DOC/AF/AF_Partie-11_Fonction_Translation_v2.3.md
   🛡️ Sécurité : instSafetyTranslationM3 (FB_Safety_Translation) câblée en parallèle
      de instTranslationM3 — SafeStop/PowerCutOff réels.
   ═══════════════════════════════════════════════════════════════ *)

PROGRAM PRG_05_Translation

VAR_INPUT
    // === 📥 ENTRÉES PROGRAMME (AUCUNE - PILOTÉ VIA PRG_02, PRG_03 & PRG_04) ===
END_VAR

VAR_OUTPUT
    // === 🚌 BUS INTER-PRG (producteur unique) ===
    Data : ST_TranslationInterPrg; // <-- [BUS] Demande finale, état public, sécurité translation M3
END_VAR

VAR
    instTranslationM3           : FB_Translation;
    instSafetyTranslationM3     : FB_Safety_Translation;
    instPosEstimatorM3          : FB_Translation_PositionEstimator;
    instOdometryGainM3          : FB_Translation_OdometryGain;    // * [INST] Gain odométrique réglable site + mesure proposée (T301)
    instPosDecoderM3            : FB_Translation_PositionDecoder; // 🧩 Decodage position M3 (migre de PRG_02, AF-02 TBD §8 #5)
    instArbM3                   : FB_TranslationCmdArbitrationM3; // * [INST] Arbitrage commande translation M3
    ArbM3_IHM                   : ST_fbTranslationCmdArbitration_IHM;     // . [LOC] Entrées IHM FB d'arbitrage M3
    ArbM3_Context               : ST_fbTranslationCmdArbitration_Context; // . [LOC] Contexte gating FB d'arbitrage M3
    ArbM3_Cfg                   : ST_fbTranslationCmdArbitration_Cfg;     // . [LOC] Config FB d'arbitrage M3 (fréquence max)

    // 🔧 Config regroupée de FB_Translation (C3 — pattern NC-110/G380, source unique GVL_PERSISTENT)
    TranslationCfg              : ST_fbTranslation_Cfg;                     // . [LOC] Cfg FB_Translation, assemblée depuis GVL_PERSISTENT

    // === 📊 STRUCTS INTERNES (publiés via Data) ===
    TranslationFinalInterlockRequest : ST_TranslationFinalInterlockRequest; // . [LOC] Demande finale et interlocks translation M3
    TranslationState                 : ST_TranslationState;                 // . [LOC] Etat public translation M3
    TranslationSafety                : ST_SafetyTranslation;                // . [LOC] Diagnostic et securites translation M3

    M3_RunRequest_Active    : BOOL;
    M3_ReqTremie_Active     : BOOL;
    M3_ReqMaintenance_Active : BOOL;
    M3_CommandConflict      : BOOL;
    M3_SpeedCmd_Active      : REAL;
    M3_PositioningActive    : BOOL;
    M3_PositionSensorTarget : BOOL;
    M3_TargetCodeSel        : INT;  // . [LOC] Code de cible M3 mémorisé (1=Trémie, 2=P2, 3=P1, 4=Maintenance) — survit à la perte de la demande
    M3_CycleTranslationStepAuthorized : BOOL; // [SAFE] En SEMI_AUTO, M3 autorise uniquement en AX2/AX14
    SimBtnIHM_Active        : BOOL; // . [LOC] Stimuli boutons IHM M3 actifs (simulation ET JoyMaster inactif)

    SelTarget       : INT;

    M3_SafeStop_Active      : BOOL; // SafeStop sur défaut module d'entrée (InputModuleFault, AF06 §3bis)
    M3_SafeStop_Aggregate   : BOOL; // 🛡️ SafeStop réellement appliqué au mouvement = InputModuleFault OR safety M3 (8 mécanismes)
    M3_MaintN2              : BOOL; // 🔒 Mode MAINT_N2 arbitré (origine FB_Modes) — garde de consommation des bypass M3

    // 🟢 Permis directionnels M3 EFFECTIFS (D1 — Phase 3) : information de POSSIBILITÉ de
    // mouvement dans une direction, donnée AVANT l'ordre. Reflète les conditions physiques/
    // logiques (fins de course, défauts, autorisation cible) — PAS la commande (homme-mort).
    // Pour M3, les conditions physiques sont calculées ici à partir des faits Safety ;
    // pas de permis secondaire (pas de benne/Kobold comme les treuils).
    EffectivePermitM3_Tremie    : BOOL; // 🟢 Permis effectif M3 vers Trémie (Safety)
    EffectivePermitM3_Maintenance : BOOL; // 🟢 Permis effectif M3 vers Maintenance (Safety)

    M3_HeightInterlockOk    : BOOL; // TRUE = M1 ET M2 au-dessus de la hauteur mini (ou bypass actif)
    M3_LimitSwitchMaintenanceEffective : BOOL; // Coupure dure §5bis — bascule sur P1 si Maintenance interdite (ex-M3_LimitSwitchRevEffective)
    M3_LimitSwitchTremieStable : BOOL; // Verrou bistable Fdc Trémie (mémorisé stable contre les rebonds) (ex-M3_LimitSwitchFwdStable)
    M3_LimitSwitchMaintenanceStable : BOOL; // Verrou bistable Fdc Maintenance/P1 (mémorisé stable contre les rebonds) (ex-M3_LimitSwitchRevStable)

    // Verrous bistables des positions cibles (§0quater) — PositionDecoder n'émet
    // plus qu'un front transitoire par capteur, mémorisé ici jusqu'à dégagement.
    M3_AtTremieStable      : BOOL;
    M3_AtPVStable          : BOOL;
    M3_AtP2Stable          : BOOL;
    M3_AtP1Stable          : BOOL;
    M3_AtMaintenanceStable : BOOL;

    // Libération du verrou §0quater sur MOUVEMENT CONFIRMÉ soutenu (fréquence réelle mesurée,
    // pas juste une consigne de sens), pendant une durée mini avant de considérer qu'on a
    // vraiment quitté le point — pas un changement de sens instantané ni un timer fixe
    // indépendant du mouvement réel (rebond capteur mal filtré).
    TonM3ConfirmedMoving : TON;
    M3_ConfirmedMoving   : BOOL;

    // FdC "soft" DIRECTIONNEL approche trémie : trémie pleine OU grille levée -> approche
    // trémie interdite, recul (Maintenance/P1) toujours libre. Distinct de la position
    // physique (M3_LimitSwitchTremieStable). PAS de latch sur recul (signal process :
    // dès qu'il retombe l'approche est re-permise). Débounce anti-parasite. Bypass N2.
    M3_TremieProcessBlock : BOOL;

    // T249-B : texte statut position M3 (lecture seule IHM) — jeton "at position" sur
    // front capteur (M3_AtXxxStable) sinon zone entre 2 capteurs (SensorsWord).
    M3_StatusText        : STRING(80);
    M3_SensorsWordPrev   : BYTE;   // detection franchissement (RAZ jeton sans dependance frequence)
    M3_SensorsWordChanged : BOOL;
    M3_AtWorkPositionStable : BOOL; // Diagnostic zone travail M3 (ne vaut pas preuve exacte d'autorisation)
    M3_AtPositionBootRestored : BOOL; // . [LOC] Restauration unique des jetons AtPosition après boot
    M3_BootRestoreApplied      : BOOL; // . [LOC] Inhibe les fronts du même scan que la restauration
    M3_BootPositionLock        : BOOL; // . [LOC] Verrou anti-RAZ des jetons pendant stabilisation boot
    M3_BootPositionLockTimer   : TON;  // . [LOC] Fenêtre de stabilisation capteurs après boot
    M3_BootSensorsWordCandidate : BYTE; // . [LOC] Mot capteurs candidat avant restauration
    M3_BootSensorsStableTimer   : TON;  // . [LOC] Validation du mot capteurs après stabilisation E/S
    TonTremieProcessBlock : TON;

    // 🕵️ Trace de blocage terrain (publiée via Data.TranslationTrace, consommée FB_TroubleshootingView)
    TranslationTrace           : ST_TraceTranslation;        // . [LOC] Trace blocage translation M3
    TraceTranslation_PrevReason : E_TranslationTraceBlockReason; // . [LOC] Cause précédente M3 (détection de changement)
END_VAR

{region "§0 Decodage position M3"}
// === 🧩 §0 DÉCODAGE POSITION M3 (migré de PRG_02, AF-02 TBD §8 #5) ===
// PRG_02_Acquisition s'exécute avant ce POU (rang 01 < 05) : HwIn.Translation est
// disponible au même scan. Le décodage des capteurs M3 est propriété de PRG_05.
instPosDecoderM3(
    SensorTremie      := PRG_02_Acquisition.HwIn.Translation.M3_PosTremie_DI,
    SensorPV          := PRG_02_Acquisition.HwIn.Translation.M3_PosPV_DI,
    SensorP2          := PRG_02_Acquisition.HwIn.Translation.M3_PosPVP2_DI,
    SensorP1          := PRG_02_Acquisition.HwIn.Translation.M3_PosP1_DI,
    SensorMaintenance := PRG_02_Acquisition.HwIn.Translation.M3_PosMaintenance_DI
);

// 📤 Publication des faits M3 dans le bus PRG_05 (consommés par PRG_07)
Data.M3_SensorWordIncoherent := instPosDecoderM3.Incoherent;
{endregion}

{region "§0 Interlock hauteur M1/M2"}
// === 🚧 §0 INTERLOCK HAUTEUR M1/M2 (risque collision translation) ===
// PRG_02_Acquisition s'exécute avant ce POU dans la MainTask (rang 01 < 05) : lecture
// du même scan, aucun retard. Bypass = maintenance consciente, doctrine ST_BypassTranslation.
// ⚠️ Une position encodeur incohérente (hors plage OU homing suspect,
// FB_Encoder_Safety) ne doit PAS pouvoir se lire comme "≥ seuil" par accident — fail-safe :
// hauteur non confirmée = interlock actif (comme une hauteur insuffisante), sauf bypass.
// 🔒 Bypass.Global NE lève PLUS cet interlock (contrairement aux autres
// causes de l'axe M3) — risque de collision jugé trop grave pour être levé par un bypass
// générique. Seul Bypass.MinHeight (dédié, conscient) lève l'anti-collision hauteur.
M3_HeightInterlockOk := GVL_IHM.M3Translation.Bypass.MinHeight
                        OR (PRG_02_Acquisition.Data.EncoderM1.HomedAndReliable
                            AND PRG_02_Acquisition.Data.EncoderM2.HomedAndReliable
                            AND (PRG_02_Acquisition.Data.EncoderM1.Measurement.CablePosM >= GVL_PERSISTENT._TranslationMinHeightM1M2_M)
                            AND (PRG_02_Acquisition.Data.EncoderM2.Measurement.CablePosM >= GVL_PERSISTENT._TranslationMinHeightM1M2_M));
TranslationState.HeightInterlockBlocking := NOT M3_HeightInterlockOk;

{endregion}

{region "§0bis Coupure dure limite translation"}
// === 🚧 §0bis COUPURE DURE (LimitSwitchMaintenance) — bascule sur P1 si Maintenance interdite ===
// LimitSwitchTremie/Maintenance protègent nativement Trémie/Maintenance
// (§5bis FB_Translation : coupure immédiate, sans rampe, dès que CommandedDirection insiste
// dans l'extrémité). P1/P2 n'ont aucune protection dure équivalente — seul le verrou souple
// (arrival-lock) les couvre. Quand Maintenance est interdite, la coupure dure doit protéger
// P1 comme si c'était l'extrémité réelle : mot 00001 (P1=0 ET Maintenance=1), UN CRAN AVANT
// la vraie extrémité Maintenance (00000) — backup si le verrou souple a déjà échoué à arrêter
// avant P1, garde la machine hors de la zone interdite plutôt que d'attendre le vrai fond.
M3_LimitSwitchMaintenanceEffective := SEL(PRG_03_Modes_Cycle.Data.Auth.MaintenanceM3TargetEnable,
                                   NOT instPosDecoderM3.TranslationPosP1 AND instPosDecoderM3.TranslationPosMaintenance,
                                   instPosDecoderM3.LimitSwitchMaintenance);

// 🔒 §0ter STABILISATION BISTABLE FINS DE COURSE EXTRÊMES (Trémie & Maintenance/P1)
// Maintient la détection stable à 1 même si le capteur physique vibre ou saute brièvement.
// Se libère uniquement sur un mouvement effectif dans le SENS INVERSE (dégagement).
// FdC LATCHE : un rebond capteur ne libere RIEN. On ne perd l'extreme Tremie qu'en
// commandant le SENS INVERSE (M3_ReqMaintenance_Active). (Ne pas rajouter de liberation
// sur mot capteurs : rebond 11111<->01111 -> flicker autorisation translation, REX MES.)
IF instPosDecoderM3.LimitSwitchTremie THEN
    M3_LimitSwitchTremieStable := TRUE;
ELSIF M3_ReqMaintenance_Active THEN
    M3_LimitSwitchTremieStable := FALSE;
END_IF;

// 🔒 §0quater FdC SOFT DIRECTIONNEL — APPROCHE TRÉMIE INTERDITE (trémie pleine / grille)
// Bloque UNIQUEMENT le sens trémie via EffectivePermitM3_Tremie ; le recul vers
// Maintenance/P1 reste libre (EffectivePermitM3_Maintenance non touché). N'entre PAS
// dans M3_LimitSwitchTremieStable -> l'info position / le voyant IHM « pont au FdC
// trémie » restent fidèles à la position physique. Aucun latch sur recul : dès que
// TremieFull_OR_GateRaised_DI retombe, l'approche est re-permise. Débounce 200 ms.
// Bypass N2 : LimitSwitch ou Global.
// ⚠️ Signal PAS ENCORE CÂBLÉ (ST_HwMachine) : polarité TRUE = bloqué à CONFIRMER au câblage.
TonTremieProcessBlock(
    IN := PRG_02_Acquisition.HwIn.Machine.TremieFull_OR_GateRaised_DI
          AND NOT GVL_IHM.M3Translation.Bypass.LimitSwitch
          AND NOT GVL_IHM.M3Translation.Bypass.Global,
    PT := T#200ms);
M3_TremieProcessBlock := TonTremieProcessBlock.Q;

// FdC LATCHE (idem Tremie) : rebond capteur ne libere rien. Perte de l'extreme
// Maintenance uniquement sur commande sens inverse (Tremie) ou sortie de la zone
// Maintenance en positionnement cible.
IF M3_LimitSwitchMaintenanceEffective THEN
    M3_LimitSwitchMaintenanceStable := TRUE;
ELSIF M3_ReqTremie_Active OR (PRG_03_Modes_Cycle.Data.Auth.MaintenanceM3TargetEnable AND NOT instPosDecoderM3.LimitSwitchMaintenance) THEN
    M3_LimitSwitchMaintenanceStable := FALSE;
END_IF;

// 🔒 §0quater MÉMORISATION DU DERNIER POINT ATTEINT (front → jeton unique)
// PositionDecoder n'émet qu'un front transitoire (1 cycle) par capteur, montant OU descendant
// SELON LE SENS (voir FB_Translation_PositionDecoder.st) — mémorisé ici pour
// tenir le niveau nécessaire au débounce (100ms) + verrou anti-rebond (§4ter DirectionAtArrival)
// de FB_Translation, et pour l'affichage IHM. MUTUELLEMENT EXCLUSIFS : un nouveau front RAZ tous
// les autres (jeton "dernier point franchi" unique). Libéré
// (RAZ complet) UNIQUEMENT sur mouvement CONFIRMÉ (fréquence réelle mesurée, pas juste la consigne
// de sens) soutenu ≥1.5s — pas un rebond capteur ni un changement de sens instantané.
M3_ConfirmedMoving := (UINT_TO_REAL(PRG_02_Acquisition.Data.M3.ActualFrequencyHz) / 100.0) > 0.5;
TonM3ConfirmedMoving(IN := M3_ConfirmedMoving, PT := T#1s500ms);

// RAZ jeton "at position" = changement du mot capteurs (franchissement reel), SANS
// dependance a la frequence variateur (souvent 0 au banc -> l'ancien RAZ ne se
// declenchait jamais -> jeton colle). Un franchissement qui EST une arrivee re-arme
// le bon jeton via les branches TranslationAtXxx ci-dessous (priorite sur la RAZ).
// Amorçage du mot précédent avant le premier calcul : un capteur déjà actif au
// boot n'est pas un franchissement et ne doit pas effacer la restauration.
IF NOT M3_AtPositionBootRestored THEN
    M3_SensorsWordPrev := instPosDecoderM3.SensorsWord;
END_IF;
M3_SensorsWordChanged := (instPosDecoderM3.SensorsWord <> M3_SensorsWordPrev);
M3_SensorsWordPrev := instPosDecoderM3.SensorsWord;
M3_BootRestoreApplied := FALSE;
M3_BootPositionLockTimer(IN := M3_BootPositionLock, PT := T#2s);
IF M3_BootPositionLock
   AND (M3_ConfirmedMoving OR M3_ReqTremie_Active OR M3_ReqMaintenance_Active OR M3_SensorsWordChanged OR M3_BootPositionLockTimer.Q) THEN
    M3_BootPositionLock := FALSE;
END_IF;

// Restauration sûre des jetons AtPosition : attendre que les E/S aient fourni
// le même mot capteurs pendant 500 ms. Sans cette attente, le premier cycle
// pouvait lire une valeur par défaut EtherCAT/CANopen (ex. P2), restaurer le
// mauvais jeton, puis verrouiller cette mauvaise position.
IF NOT M3_AtPositionBootRestored THEN
    IF instPosDecoderM3.SensorsWord <> M3_BootSensorsWordCandidate THEN
        M3_BootSensorsWordCandidate := instPosDecoderM3.SensorsWord;
        M3_BootSensorsStableTimer(IN := FALSE, PT := T#500ms);
    ELSE
        M3_BootSensorsStableTimer(IN := TRUE, PT := T#500ms);
    END_IF;
ELSE
    M3_BootSensorsStableTimer(IN := FALSE, PT := T#500ms);
END_IF;

// Le RETAIN n'est accepté que si le mot capteurs présent au boot est stable.
// Si le pont a bougé hors tension, aucun ancien jeton n'est réinjecté.
IF NOT M3_AtPositionBootRestored
   AND NOT M3_ConfirmedMoving
   AND NOT M3_ReqTremie_Active
   AND NOT M3_ReqMaintenance_Active
   AND M3_BootSensorsStableTimer.Q THEN
    CASE instPosDecoderM3.SensorsWord OF
        2#11111:
            M3_AtTremieStable := GVL_PERSISTENT._TranslationAtTremiePersisted OR instPosDecoderM3.TranslationPosTremie;
            M3_AtPVStable := FALSE; M3_AtP2Stable := FALSE; M3_AtP1Stable := FALSE; M3_AtMaintenanceStable := FALSE;
        2#01111:
            M3_AtPVStable := GVL_PERSISTENT._TranslationAtPVPersisted OR instPosDecoderM3.TranslationPosPV;
            M3_AtTremieStable := FALSE; M3_AtP2Stable := FALSE; M3_AtP1Stable := FALSE; M3_AtMaintenanceStable := FALSE;
        2#00111:
            M3_AtP2Stable := GVL_PERSISTENT._TranslationAtP2Persisted OR instPosDecoderM3.TranslationPosP2;
            M3_AtTremieStable := FALSE; M3_AtPVStable := FALSE; M3_AtP1Stable := FALSE; M3_AtMaintenanceStable := FALSE;
        2#00011:
            M3_AtP1Stable := GVL_PERSISTENT._TranslationAtP1Persisted OR instPosDecoderM3.TranslationPosP1;
            M3_AtTremieStable := FALSE; M3_AtPVStable := FALSE; M3_AtP2Stable := FALSE; M3_AtMaintenanceStable := FALSE;
        2#00000:
            M3_AtMaintenanceStable := GVL_PERSISTENT._TranslationAtMaintenancePersisted OR instPosDecoderM3.TranslationPosMaintenance;
            M3_AtTremieStable := FALSE; M3_AtPVStable := FALSE; M3_AtP2Stable := FALSE; M3_AtP1Stable := FALSE;
    END_CASE;
    M3_AtPositionBootRestored := TRUE;
    M3_BootRestoreApplied := TRUE;
    M3_BootPositionLock := TRUE;
END_IF;

IF NOT M3_BootPositionLock AND NOT M3_BootRestoreApplied AND instPosDecoderM3.TranslationAtTremie THEN
    M3_AtTremieStable := TRUE; M3_AtPVStable := FALSE; M3_AtP2Stable := FALSE; M3_AtP1Stable := FALSE; M3_AtMaintenanceStable := FALSE;
ELSIF NOT M3_BootPositionLock AND NOT M3_BootRestoreApplied AND instPosDecoderM3.TranslationAtPV THEN
    M3_AtPVStable := TRUE; M3_AtTremieStable := FALSE; M3_AtP2Stable := FALSE; M3_AtP1Stable := FALSE; M3_AtMaintenanceStable := FALSE;
ELSIF NOT M3_BootPositionLock AND NOT M3_BootRestoreApplied AND instPosDecoderM3.TranslationAtP2 THEN
    M3_AtP2Stable := TRUE; M3_AtTremieStable := FALSE; M3_AtPVStable := FALSE; M3_AtP1Stable := FALSE; M3_AtMaintenanceStable := FALSE;
ELSIF NOT M3_BootPositionLock AND NOT M3_BootRestoreApplied AND instPosDecoderM3.TranslationAtP1 THEN
    M3_AtP1Stable := TRUE; M3_AtTremieStable := FALSE; M3_AtPVStable := FALSE; M3_AtP2Stable := FALSE; M3_AtMaintenanceStable := FALSE;
ELSIF NOT M3_BootPositionLock AND NOT M3_BootRestoreApplied AND instPosDecoderM3.TranslationAtMaintenance THEN
    M3_AtMaintenanceStable := TRUE; M3_AtTremieStable := FALSE; M3_AtPVStable := FALSE; M3_AtP2Stable := FALSE; M3_AtP1Stable := FALSE;
ELSIF NOT M3_BootPositionLock AND NOT M3_BootRestoreApplied AND M3_SensorsWordChanged THEN
    // Le mot capteurs a change sans que ce soit une arrivee -> on a quitte le dernier point.
    // Tremie/Maintenance EXCLUS ICI (rebond capteur) : ils suivent desormais la regle
    // bistable ci-dessous, identique et deja prouvee sur LimitSwitchTremie/MaintenanceStable §0ter.
    M3_AtPVStable := FALSE; M3_AtP2Stable := FALSE; M3_AtP1Stable := FALSE;
END_IF;

// Bistable Tremie/Maintenance : jamais efface par un rebond capteur (mot capteurs),
// uniquement par une commande franche dans le sens inverse — meme regle, deja prouvee
// sans regression depuis 2026-09-04, que M3_LimitSwitchTremieStable/MaintenanceStable §0ter.
IF M3_ReqMaintenance_Active THEN
    M3_AtTremieStable := FALSE;
END_IF;
IF GVL_IHM.M3Translation.Cmd.BtnSetAtP1 THEN
    M3_AtP1Stable := TRUE;
    M3_AtTremieStable := FALSE;
    M3_AtPVStable := FALSE;
    M3_AtP2Stable := FALSE;
    M3_AtMaintenanceStable := FALSE;
END_IF;
IF M3_ReqTremie_Active THEN
    M3_AtMaintenanceStable := FALSE;
END_IF;

// --- M3 a une position de travail : STATIQUE (mot capteurs), pas un jeton de franchissement ---
// Les jetons M3_AtXxxStable ne se posent que sur un FRONT capteur : au boot PLC, pont deja
// pose a P1 ou Maintenance sans mouvement -> jetons FALSE -> le verrou descente treuil
// (T249-A) resterait bloque jusqu'a devoir franchir un capteur. On complete donc par une
// lecture STATIQUE du mot : 00011 = zone P2->P1 (capteur P1 fait, P2 depasse) ; 00000 =
// extreme Maintenance.
// ATTENTION : 00011 couvre TOUTE la zone P2->P1 (15..20 m), pas le seul point P1. On
// n'autorise donc la lecture statique QUE si le pont est A L'ARRET et sans cible en cours,
// sinon la descente treuil serait permise pendant le transit P2->P1 (5 m). Le jeton
// M3_AtP1Stable (front) reste la voie normale quand le pont vient d'arriver.
// Information de supervision uniquement : 00011 couvre toute la zone P2->P1.
// Le verrou de descente consomme directement les jetons AtP1/AtMaintenance.
M3_AtWorkPositionStable := (NOT instPosDecoderM3.Incoherent)
    AND ( M3_AtP1Stable OR M3_AtMaintenanceStable
          OR ( (instPosDecoderM3.SensorsWord = 2#00011 OR instPosDecoderM3.SensorsWord = 2#00000)
               AND NOT M3_ConfirmedMoving
               AND NOT M3_ReqTremie_Active
               AND NOT M3_ReqMaintenance_Active ) );

// Mémorisation persistante : un mot capteurs exact et stable au repos prime
// sur le jeton RAM, qui peut avoir été perdu juste avant la coupure.
IF NOT M3_ConfirmedMoving
   AND NOT M3_ReqTremie_Active
   AND NOT M3_ReqMaintenance_Active THEN
    CASE instPosDecoderM3.SensorsWord OF
        2#11111:
            GVL_PERSISTENT._TranslationAtTremiePersisted := TRUE;
            GVL_PERSISTENT._TranslationAtPVPersisted := FALSE;
            GVL_PERSISTENT._TranslationAtP2Persisted := FALSE;
            GVL_PERSISTENT._TranslationAtP1Persisted := FALSE;
            GVL_PERSISTENT._TranslationAtMaintenancePersisted := FALSE;
        2#01111:
            GVL_PERSISTENT._TranslationAtTremiePersisted := FALSE;
            GVL_PERSISTENT._TranslationAtPVPersisted := TRUE;
            GVL_PERSISTENT._TranslationAtP2Persisted := FALSE;
            GVL_PERSISTENT._TranslationAtP1Persisted := FALSE;
            GVL_PERSISTENT._TranslationAtMaintenancePersisted := FALSE;
        2#00111:
            GVL_PERSISTENT._TranslationAtTremiePersisted := FALSE;
            GVL_PERSISTENT._TranslationAtPVPersisted := FALSE;
            GVL_PERSISTENT._TranslationAtP2Persisted := TRUE;
            GVL_PERSISTENT._TranslationAtP1Persisted := FALSE;
            GVL_PERSISTENT._TranslationAtMaintenancePersisted := FALSE;
        2#00011:
            GVL_PERSISTENT._TranslationAtTremiePersisted := FALSE;
            GVL_PERSISTENT._TranslationAtPVPersisted := FALSE;
            GVL_PERSISTENT._TranslationAtP2Persisted := FALSE;
            GVL_PERSISTENT._TranslationAtP1Persisted := TRUE;
            GVL_PERSISTENT._TranslationAtMaintenancePersisted := FALSE;
        2#00000:
            GVL_PERSISTENT._TranslationAtTremiePersisted := FALSE;
            GVL_PERSISTENT._TranslationAtPVPersisted := FALSE;
            GVL_PERSISTENT._TranslationAtP2Persisted := FALSE;
            GVL_PERSISTENT._TranslationAtP1Persisted := FALSE;
            GVL_PERSISTENT._TranslationAtMaintenancePersisted := TRUE;
        ELSE
            GVL_PERSISTENT._TranslationAtTremiePersisted := M3_AtTremieStable;
            GVL_PERSISTENT._TranslationAtPVPersisted := M3_AtPVStable;
            GVL_PERSISTENT._TranslationAtP2Persisted := M3_AtP2Stable;
            GVL_PERSISTENT._TranslationAtP1Persisted := M3_AtP1Stable;
            GVL_PERSISTENT._TranslationAtMaintenancePersisted := M3_AtMaintenanceStable;
    END_CASE;
END_IF;

{endregion}

{region "§1 Arbitrage cible et direction"}
// === 🔀 §1 ARBITRAGE DU SÉLECTEUR DE CIBLE ET DE LA DIRECTION ===

// ── Arbitrage M3 (FB_TranslationCmdArbitrationM3) ──
// Remplissage des structs d'arbitrage (champ par champ, CODESYS 3.5 refuse l'init anonyme en appel)
// 🎛️ Stimuli boutons IHM M3 : en simulation ET JoyMaster inactif, les stimuli pilotent les
// boutons IHM (SEL) ; sinon la valeur IHM réelle est conservée (jamais écrasée, producteur unique).
SimBtnIHM_Active := GVL_Simulation.SimulationModeActive AND NOT GVL_IHM.Modes.Cmd.TglJoystickMaster;
ArbM3_IHM.BtnTremie         := SEL(SimBtnIHM_Active, GVL_IHM.M3Translation.Cmd.BtnTremie, GVL_Simulation.SimBtnTremie);
ArbM3_IHM.BtnMaintenance    := SEL(SimBtnIHM_Active, GVL_IHM.M3Translation.Cmd.BtnMaintenance, GVL_Simulation.SimBtnMaintenance);
ArbM3_IHM.SelPositioning    := GVL_IHM.M3Translation.Cmd.SelPositioning;
ArbM3_IHM.SetFreq_Hz        := GVL_IHM.M3Translation.Cmd.SetFreq_Hz;
ArbM3_IHM.BypassGlobal      := GVL_IHM.M3Translation.Bypass.Global;

ArbM3_Context.HeightInterlockOk := M3_HeightInterlockOk;
ArbM3_Cfg.MaxFreq_Hz            := GVL_PERSISTENT._TranslationMaxFreq_Hz;

instArbM3(
    Enable         := TRUE,
    Joystick       := PRG_02_Acquisition.Data.Joystick,
    Auth           := PRG_03_Modes_Cycle.Data.Auth,
    ReqTranslation := PRG_03_Modes_Cycle.Data.ReqProgram.ReqTranslation,
    IHM            := ArbM3_IHM,
    TglJoystickMaster := GVL_IHM.Modes.Cmd.TglJoystickMaster,
    Context        := ArbM3_Context,
    Cfg            := ArbM3_Cfg
);
M3_PositioningActive := instArbM3.PositioningActive;
SelTarget := instArbM3.SelTarget;
M3_RunRequest_Active := instArbM3.RunRequest;
M3_ReqTremie_Active := instArbM3.ReqTremie;
M3_ReqMaintenance_Active := instArbM3.ReqMaintenance;
M3_CommandConflict := instArbM3.CommandConflict;
M3_SpeedCmd_Active := instArbM3.SpeedPct;

// Verrou independant du G7 et de l'arbitrage joystick : en SEMI_AUTO, aucune
// commande M3 ne doit survivre hors des deux etapes explicitement dediees a la
// translation. Ce veto couvre notamment AX3/AX10/AX15 (manoeuvres benne), meme
// si une demande ReqTranslation ou un etat interne restait accidentellement actif.
M3_CycleTranslationStepAuthorized :=
    (PRG_03_Modes_Cycle.Data.SequenceState.Step = E_AutoCycleStep.AX2_TRANSLATE_P1)
    OR (PRG_03_Modes_Cycle.Data.SequenceState.Step = E_AutoCycleStep.AX14_TRANSLATE_DUMP);

IF (PRG_03_Modes_Cycle.Data.Auth.Mode = E_Mode.SEMI_AUTO)
   AND NOT M3_CycleTranslationStepAuthorized THEN
    M3_RunRequest_Active := FALSE;
    M3_ReqTremie_Active := FALSE;
    M3_ReqMaintenance_Active := FALSE;
    M3_SpeedCmd_Active := 0.0;
END_IF;

// InvertDirection est appliqué dans FB_Translation (InvertDriveDirection), uniquement au mot
// de commande variateur en sortie — les bits ReqTremie/ReqMaintenance restent le sens sémantique réel.

// 🩺 InputModuleFault (AF06 §3bis) : un module DI TOR hors service rend indisponibles
// les retours frein/thermique/positions du VH_0808ETP/VH_0800END portant M3 — rampe rapide.
M3_SafeStop_Active := PRG_02_Acquisition.Data.InputModules.Fault;

// En mode manuel (SelTarget=0), n'importe quel des 3 points d'arrêt (Trémie/P1/Maintenance)
// arme le verrou anti-rebond §4ter de FB_Translation (DirectionAtArrival). Mot EXACT
// (TranslationAtXxx), pas le cumulatif (TranslationPosXxx) — front franc à l'arrivée quel que
// soit le sens de venue (voir FB_Translation_PositionDecoder.st).
//
// 🎯 MÉMOIRE DE CIBLE : le code de cible n'est réécrit QUE tant qu'une demande est présente ;
// la cible publiée est ensuite le JETON du point mémorisé. La perte de la demande n'efface donc
// plus une cible déjà qualifiée : le debounce de 100 ms de FB_Translation peut se terminer et
// armer son verrou d'arrivée même si l'opérateur relâche juste après le capteur. Sans cette
// mémoire, un relâchement dans la fenêtre de debounce annulait la détection d'arrivée en cours,
// et la re-demande du même sens repartait au-delà du point. La cible retombe d'elle-même dès que
// le chariot quitte le point, les jetons M3_AtXxxStable étant uniques et exclusifs.
// La voie directionnelle reste celle du mode manuel : en SEMI_AUTO la cible d'étape est fournie
// par SelTarget (1 en AX14, 3 en AX2) et ne dépend d'aucune demande.
CASE SelTarget OF
    1: M3_TargetCodeSel := 1;
    2: M3_TargetCodeSel := 2;
    3: M3_TargetCodeSel := 3;
    4: M3_TargetCodeSel := 4;
ELSE
    IF M3_ReqTremie_Active THEN
        // En Marche Avant (+1 vers Trémie) : seule Trémie est le point d'arrêt automatique
        M3_TargetCodeSel := 1;
    ELSIF M3_ReqMaintenance_Active THEN
        // En Marche Arrière (-1 vers Maintenance) :
        // - Si Maintenance autorisée -> arrêt sur Maintenance
        // - Si Maintenance interdite -> arrêt sur P1
        IF PRG_03_Modes_Cycle.Data.Auth.MaintenanceM3TargetEnable THEN
            M3_TargetCodeSel := 4;
        ELSE
            M3_TargetCodeSel := 3;
        END_IF;
    END_IF;
END_CASE;

CASE M3_TargetCodeSel OF
    1: M3_PositionSensorTarget := M3_AtTremieStable;
    2: M3_PositionSensorTarget := M3_AtP2Stable;
    3: M3_PositionSensorTarget := M3_AtP1Stable;
    4: M3_PositionSensorTarget := M3_AtMaintenanceStable;
ELSE
    M3_PositionSensorTarget := FALSE;
END_CASE;

{endregion}

{region "§1bis Garde de mode des bypass M3"}
// 🔒 Les bypass de l'axe M3 sont actionnables UNIQUEMENT en MAINT_N2 (doctrine
// ST_BypassTranslation.st) : le bit RETAIN restauré au boot est sinon consommé sans aucune
// garde de mode. Un seul bit de fin de course neutralise TROIS barrières de l'axe — le verrou
// d'arrivée et la cause 6 de FB_Translation, et la cause 6 de FB_Safety_Translation — soit la
// neutralisation des sécurités de fin de course depuis un mode de marche nominal.
// La garde est posée AU POINT DE CONSOMMATION : le stockage RETAIN et sa restauration vers
// l'IHM ne sont pas touchés, le bit reste donc lisible et actionnable en MAINT_N2.
// Origine du mode = arbitrage FB_Modes (Auth.Mode), jamais le sélecteur IHM brut — même
// exigence que la garde des bypass treuils.
M3_MaintN2 := (PRG_03_Modes_Cycle.Data.Auth.Mode = E_Mode.MAINT_N2);
{endregion}

{region "§1bis Securite M3"}
// === 🛡️ §1bis SÉCURITÉ M3 (FB_Safety_Translation, câblée en parallèle visible) ===
// ⚠️ Ordre d'appel volontaire : la safety lit ici le BrakeReleaseRequest et le
// BrakeCmd du SCAN PRÉCÉDENT d'instTranslationM3 (elle est appelée avant), soit un retard
// d'un scan. Bénin : BrakeReleaseRequest ne change pas plus vite qu'un scan MainTask 10 ms
// sur une commande frein.
instSafetyTranslationM3(
    Enable                  := (PRG_03_Modes_Cycle.Data.Auth.Mode <> E_Mode.DISABLE),
    Reset                   := PRG_07_Supervision.FaultMachineReset_IHM,
    PowerContactorEngaged   := PRG_02_Acquisition.HwIn.Machine.PowerContactorEngaged_DI,
    Mode                    := PRG_03_Modes_Cycle.Data.Auth.Mode,
    JoystickOnline          := PRG_02_Acquisition.Data.Network.Joystick.Online,
    JoystickOperational     := PRG_02_Acquisition.Data.Network.Joystick.Operational,
    HeartbeatIhmOk          := GVL_IHM.Commun.HeartbeatIhmOk,
    PhaseRotationOk         := PRG_02_Acquisition.HwIn.Machine.PhaseRotationOk_DI,
    BrakeThermalFeedback    := NOT PRG_02_Acquisition.HwIn.Machine.M1_M2_M3_BrakeThermalOk_DI,
    DriveOnline             := PRG_02_Acquisition.Data.Network.DriveM3.Online,
    DriveOperational        := PRG_02_Acquisition.Data.Network.DriveM3.Operational,
    DriveStatusWord         := PRG_02_Acquisition.Data.M3.StatusWord,
    DriveActualFreqHz       := UINT_TO_REAL(PRG_02_Acquisition.Data.M3.ActualFrequencyHz) / 100.0,
    BrakeFeedback           := SEL(GVL_IHM.M3Translation.Bypass.ContactorFeedback OR GVL_IHM.M3Translation.Bypass.Global, PRG_02_Acquisition.HwIn.Translation.M3_BrakeIsOpen_DI, instTranslationM3.BrakeReleaseRequest),
    BrakeCmd                := instTranslationM3.BrakeReleaseRequest,
    RunRequest              := M3_RunRequest_Active,
    ReqTremie               := M3_ReqTremie_Active,
    ReqMaintenance          := M3_ReqMaintenance_Active,
    LimitSwitchTremie       := M3_LimitSwitchTremieStable,
    LimitSwitchMaintenance  := M3_LimitSwitchMaintenanceStable,
    SensorWordIncoherent    := instPosDecoderM3.Incoherent,
    BypassGlobal            := GVL_IHM.M3Translation.Bypass.Global,
    BypassOperatorComm      := GVL_IHM.M3Translation.Bypass.OperatorComm,
    BypassDriveComm         := GVL_IHM.M3Translation.Bypass.DriveComm,
    BypassPhaseRotation     := GVL_IHM.M3Translation.Bypass.PhaseRotation,
    BypassBrakeThermal      := GVL_IHM.M3Translation.Bypass.BrakeThermal,
    BypassMecaB             := GVL_IHM.M3Translation.Bypass.MecaB,
    BypassMecaA             := GVL_IHM.M3Translation.Bypass.MecaA,
    BypassLimitSwitch       := M3_MaintN2 AND (GVL_IHM.M3Translation.Bypass.LimitSwitch OR GVL_IHM.M3Translation.Bypass.Global),
    BypassSensorIncoherent  := GVL_IHM.M3Translation.Bypass.SensorIncoherent,
    BypassSafety            := GVL_IHM.M3Translation.Bypass.Safety,
    BypassProcess           := GVL_IHM.M3Translation.Bypass.Process
);

// SafeStop réellement appliqué au mouvement = agrégat InputModuleFault OR safety M3
// (8 mécanismes) — aucune des deux causes ne doit être perdue.
// + Verrou translation pendant le cycle de homing machine (HX2..HX6) : le chariot M3
//   ne doit pas bouger tant que M1/M2 se référencent (produit par FB_CycleMachineHoming,
//   publié PRG_02.Data.MachineHoming.M3Locked). Pas de bypass : conscient = quitter le cycle.
M3_SafeStop_Aggregate := M3_SafeStop_Active
                         OR instSafetyTranslationM3.SafeStop
                         OR PRG_02_Acquisition.Data.MachineHoming.M3Locked;

{endregion}

{region "§1ter Permis effectifs M3 (D1)"}
// === 🟢 §1ter PERMIS EFFECTIFS M3 (D1 — Phase 3) ===
// Niveau exposé à l'IHM = EFFECTIF, aligné sur les treuils M1/M2 (PRG_04 §5).
// ⚠️ Le permit est une INFORMATION DE POSSIBILITÉ de mouvement dans une direction,
// donnée AVANT l'ordre. Il reflète que l'axe est PRÊT À FONCTIONNER (pas de défaut,
// puissance, thermique) ET que la direction est physiquement possible (fins de course,
// autorisation cible). Il ne reflète PAS la commande (homme-mort) : l'homme-mort est une
// condition de COMMANDE (arbitrage FB_TranslationCmdArbitrationM3 / FB_CycleSemiAuto), pas de
// possibilité — il n'entre donc PAS dans le permit exposé.
// Pour M3, le Safety (FB_Safety_Translation) fournit les faits de sécurité :
//   - TremieLimitClear = NOT LimitSwitchTremie (direction possible vers Trémie)
//   - MaintenanceLimitClear = NOT LimitSwitchMaintenance (direction possible jusqu'à P1)
//   - SafeStop / PowerCutOff = défauts (thermique, Méca A/B, incohérence, comm, phases...)
// Le permis effectif = fait de limite libre AND NOT SafeStop AND NOT PowerCutOff
// (prêt à fonctionner), aligné sur le modèle treuils où le Safety produit déjà des
// permis gatés par les défauts. Pas de Process supplémentaire (pas de benne/Kobold).
// ⚠️ Le verrou « descente treuil interdite tant que M3 pas à P1 » (DumpAtTremieDescentLocked)
// est côté TREUIL (PRG_04 §5, lignes 802-805), pas dans le permit M3 : le permit M3 reste une
// information de possibilité de mouvement de la translation, indépendante de l'état de la trémie.
// ⚠️ Le permit M3 est un permit EFFECTIF « pouvoir bouger » (prêt à fonctionner), PAS un pur
// directionnel. Quand l'axe est en défaut (SafeStop/PowerCutOff), TOUS les sens sont bloqués ;
// au retour en condition, un sens peut être permis et pas l'autre. L'interdiction d'accès à la
// zone Maintenance ne retire PAS le permis de rejoindre P1 : elle agit sur la cible et la
// coupure dure M3_LimitSwitchMaintenanceEffective.
EffectivePermitM3_Tremie    := instSafetyTranslationM3.TremieLimitClear
                               AND NOT M3_SafeStop_Aggregate
                               AND NOT instSafetyTranslationM3.PowerCutOff
                               AND NOT M3_TremieProcessBlock;
EffectivePermitM3_Maintenance := instSafetyTranslationM3.MaintenanceLimitClear
                                  AND NOT M3_SafeStop_Aggregate
                                  AND NOT instSafetyTranslationM3.PowerCutOff;

{endregion}

{region "§2 Pilotage translation M3"}
// === ⚙️ §2 EXÉCUTION PILOTAGE TRANSLATION M3 ===

// 🔧 Assemblage de la config FB_Translation (C3) — SOURCE UNIQUE : GVL_PERSISTENT.
// Fini le double sourcing (rampes flat + vitesses d'approche via GVL_IHM.M3Translation.Cfg).
// Les 3 vitesses d'approche sont lues dans _TranslationCfgPersist (miroir persistant de
// ST_TranslationCfg, synchronisé par FB_CfgPersistBridge_TranslationCfg dans PRG_07) — la
// valeur reflète toute modification IHM persistée. Les délais (DirectionInterlockDelay,
// CaptorDebounce, BrakeDelay*, BrakeFeedbackTimeout) restent aux valeurs défaut du struct
// (non réglés IHM) — même comportement qu'avant (non câblés, défauts FB).
TranslationCfg.CfgRampAccelRate           := _TranslationRampAccelRate_Pct;
TranslationCfg.CfgRampDecelNormalRate     := _TranslationRampDecelNormal_Pct;
TranslationCfg.CfgRampDecelFastRate       := _TranslationRampDecelFast_Pct;
TranslationCfg.DriveFreqScaleMaxHz        := _TranslationMaxFreq_Hz;
TranslationCfg.ApproachSpeedTremieHz      := _TranslationCfgPersist.CfgApproachSpeedTremie_Hz;
TranslationCfg.ApproachSpeedMaintenanceHz := _TranslationCfgPersist.CfgApproachSpeedMaintenance_Hz;
TranslationCfg.ApproachSpeedP1Hz          := _TranslationCfgPersist.CfgApproachSpeedP1_Hz;

instTranslationM3(
    Enable                  := (PRG_03_Modes_Cycle.Data.Auth.Mode <> E_Mode.DISABLE),
    Reset                   := PRG_07_Supervision.FaultMachineReset_IHM,
    PowerContactorEngaged   := PRG_02_Acquisition.HwIn.Machine.PowerContactorEngaged_DI,
    Mode                    := PRG_03_Modes_Cycle.Data.Auth.Mode,
    RunRequest              := M3_RunRequest_Active,
    SafeStop                := M3_SafeStop_Aggregate,
    ReqTremie               := M3_ReqTremie_Active,
    ReqMaintenance          := M3_ReqMaintenance_Active,
    InvertDriveDirection    := GVL_IHM.M3Translation.Cmd.InvertDirection,
    SpeedTgt_Pct            := M3_SpeedCmd_Active,
    PositionSensorTarget    := M3_PositionSensorTarget,
    SlowdownSensorTremie       := instPosDecoderM3.TranslationPosPV,
    // Les 5 capteurs forment un code thermomètre cumulatif depuis la Trémie (voir
    // FB_Translation_PositionDecoder.st). Chaque zone est délimitée par "capteur PRÉCÉDENT retombé
    // à 0" ET "capteur de la zone encore à 1" — zone P2→P1 = NOT PosP2 AND PosP1 (mot 00011) ;
    // zone P1→Maintenance = NOT PosP1 AND PosMaintenance (mot 00001). Zones mutuellement exclusives,
    // chacune sa propre vitesse d'approche (CfgApproachSpeedP1_Hz / CfgApproachSpeedMaintenance_Hz).
    SlowdownSensorMaintenance  := (NOT instPosDecoderM3.TranslationPosP1) AND instPosDecoderM3.TranslationPosMaintenance,
    // Ralentissement P2→P1 UNIQUEMENT si P1 est un vrai point
    // d'arrêt (zone Maintenance NON autorisée). Zone Maintenance autorisée -> 100% vitesse jusqu'à
    // P1, ralentissement seulement après (zone P1→Maintenance, SlowdownSensorMaintenance ci-dessus).
    SlowdownSensorP1           := (NOT instPosDecoderM3.TranslationPosP2) AND instPosDecoderM3.TranslationPosP1
                                   AND NOT PRG_03_Modes_Cycle.Data.Auth.MaintenanceM3TargetEnable,
    LimitSwitchTremie       := M3_LimitSwitchTremieStable,
    LimitSwitchMaintenance  := M3_LimitSwitchMaintenanceStable,
    // 🛡️ Permis directionnels SAFETY (source unique instSafetyTranslationM3) — gate de sens FB_Translation
    EffectivePermitM3_Tremie := EffectivePermitM3_Tremie,
    EffectivePermitM3_Maintenance := EffectivePermitM3_Maintenance,
    DriveStatusWord         := PRG_02_Acquisition.Data.M3.StatusWord,
    DriveActualFreqHz       := UINT_TO_REAL(PRG_02_Acquisition.Data.M3.ActualFrequencyHz) / 100.0,
    Cfg                     := TranslationCfg,
    BrakeFeedback           := SEL(GVL_IHM.M3Translation.Bypass.ContactorFeedback OR GVL_IHM.M3Translation.Bypass.Global, PRG_02_Acquisition.HwIn.Translation.M3_BrakeIsOpen_DI, instTranslationM3.BrakeReleaseRequest),
    BypassContactorCheck    := GVL_IHM.M3Translation.Bypass.Global OR GVL_IHM.M3Translation.Bypass.ContactorFeedback,
    BypassLimitSwitch       := M3_MaintN2 AND (GVL_IHM.M3Translation.Bypass.Global OR GVL_IHM.M3Translation.Bypass.LimitSwitch)
);

// 📏 Gain odométrique (T301) : réglage site |P2-PV| / (CalibFreq × CalibTime), repli sur le gain
// persistant si non saisi. La mesure P2 <-> PV est PROPOSÉE (State.OdometryMeasured*), jamais appliquée.
instOdometryGainM3(
    Enable               := (PRG_03_Modes_Cycle.Data.Auth.Mode <> E_Mode.DISABLE),
    SensorPV             := instPosDecoderM3.TranslationPosPV,
    SensorP2             := instPosDecoderM3.TranslationPosP2,
    DriveActualFreq_Hz   := TO_REAL(PRG_02_Acquisition.Data.M3.ActualFrequencyHz) / 100.0,
    PosPV_M              := GVL_PERSISTENT._TranslationPosPV_M,
    PosP2_M              := GVL_PERSISTENT._TranslationPosP2_M,
    CalibFreq_Hz         := GVL_PERSISTENT._TranslationCalibFreq_Hz,
    CalibTime_S          := GVL_PERSISTENT._TranslationCalibTimeP2PV_S,
    FallbackGain         := GVL_PERSISTENT._TranslationGainMetersPerHzSec
);

// 📐 Estimateur de position continue M3 (odométrie + recalage 5 capteurs)
instPosEstimatorM3(
    Enable               := (PRG_03_Modes_Cycle.Data.Auth.Mode <> E_Mode.DISABLE),
    Reset                := PRG_07_Supervision.FaultMachineReset_IHM,
    DriveActualFreqHz    := TO_REAL(PRG_02_Acquisition.Data.M3.ActualFrequencyHz) / 100.0,
    ReqTremie            := M3_ReqTremie_Active,
    ReqMaintenance       := M3_ReqMaintenance_Active,
    SensorMaintenance    := instPosDecoderM3.TranslationPosMaintenance,
    SensorP1             := instPosDecoderM3.TranslationPosP1,
    SensorP2             := instPosDecoderM3.TranslationPosP2,
    SensorPV             := instPosDecoderM3.TranslationPosPV,
    SensorTremie         := instPosDecoderM3.TranslationPosTremie,
    PosMaintenanceM      := GVL_PERSISTENT._TranslationPosMaintenance_M,
    PosP1M               := GVL_PERSISTENT._TranslationPosP1_M,
    PosP2M               := GVL_PERSISTENT._TranslationPosP2_M,
    PosPVM               := GVL_PERSISTENT._TranslationPosPV_M,
    PosTremieM           := GVL_PERSISTENT._TranslationPosTremie_M,
    GainMetersPerHzSec   := instOdometryGainM3.GainActive,
    PersistedPositionM   := GVL_PERSISTENT._TranslationPosEstimated_M,
    PersistedInitialized := GVL_PERSISTENT._TranslationPosEstimatedInitialized
);
// Recopie continue (reprise après reboot, doctrine _TranslationSetFreq_Hz) — pas de bridge dédié.
GVL_PERSISTENT._TranslationPosEstimated_M := instPosEstimatorM3.PositionEstimatedM;
GVL_PERSISTENT._TranslationPosEstimatedInitialized := instPosEstimatorM3.Initialized;

// === T249-B : TEXTE STATUT POSITION M3 (lecture seule IHM) ============================
// Source = jeton "at position" sur front capteur (M3_AtXxxStable, mecanisme d'origine,
// RAZ sur changement de mot capteurs). Sinon zone entre 2 capteurs via SensorsWord
// (code thermometre cumulatif). AUCUNE dependance a la frequence variateur.
IF M3_AtTremieStable THEN
    M3_StatusText := 'M3 a la Tremie';
ELSIF M3_AtMaintenanceStable THEN
    M3_StatusText := 'M3 a la Maintenance';
ELSIF M3_AtP1Stable THEN
    M3_StatusText := 'M3 a P1';
ELSIF M3_AtP2Stable THEN
    M3_StatusText := 'M3 a P2';
ELSIF M3_AtPVStable THEN
    M3_StatusText := 'M3 a PV';
ELSIF instPosDecoderM3.Incoherent THEN
    M3_StatusText := 'M3 capteurs INCOHERENTS';
ELSE
    CASE instPosDecoderM3.SensorsWord OF
        2#11111: M3_StatusText := 'M3 a la Tremie';
        2#01111: M3_StatusText := 'M3 entre Tremie et PV';
        2#00111: M3_StatusText := 'M3 entre PV et P2';
        2#00011: M3_StatusText := 'M3 entre P2 et P1';
        2#00001: M3_StatusText := 'M3 entre P1 et Maintenance';
        2#00000: M3_StatusText := 'M3 a la Maintenance';
    ELSE
        M3_StatusText := 'M3 position indeterminee';
    END_CASE;
END_IF;
// Suffixe sens de deplacement (commande active).
IF M3_ReqTremie_Active THEN
    M3_StatusText := CONCAT(M3_StatusText, ' -> Tremie');
ELSIF M3_ReqMaintenance_Active THEN
    M3_StatusText := CONCAT(M3_StatusText, ' -> Maintenance');
END_IF;

{endregion}

{region "§3 Publication demande translation"}
// === 📤 §3 PUBLICATION DEMANDE BRUTE TRANSLATION ===

TranslationFinalInterlockRequest.Enable := (PRG_03_Modes_Cycle.Data.Auth.Mode <> E_Mode.DISABLE);
TranslationFinalInterlockRequest.Reset := PRG_07_Supervision.FaultMachineReset_IHM;
TranslationFinalInterlockRequest.PowerContactorEngaged := PRG_02_Acquisition.HwIn.Machine.PowerContactorEngaged_DI;
TranslationFinalInterlockRequest.SafeStop := M3_SafeStop_Aggregate;
TranslationFinalInterlockRequest.PowerCutOff := instSafetyTranslationM3.PowerCutOff;
TranslationFinalInterlockRequest.EffectivePermitM3_Tremie := EffectivePermitM3_Tremie;
TranslationFinalInterlockRequest.EffectivePermitM3_Maintenance := EffectivePermitM3_Maintenance;
TranslationFinalInterlockRequest.BrakeReleaseRequest := instTranslationM3.BrakeReleaseRequest;
TranslationFinalInterlockRequest.BrakeCommandOpenConfirmed := instTranslationM3.BrakeCommandOpenConfirmed;
TranslationFinalInterlockRequest.RequestedDriveControlWord := instTranslationM3.RequestedDriveControlWord;
TranslationFinalInterlockRequest.RequestedDriveFreqHz := instTranslationM3.RequestedDriveFreqHz;
TranslationFinalInterlockRequest.ReqTremieSemantic := M3_ReqTremie_Active;
TranslationFinalInterlockRequest.ReqMaintenanceSemantic := M3_ReqMaintenance_Active;

// Derniere barriere avant PRG_06 : neutralisation immediate du variateur ET du
// frein M3 hors AX2/AX14 en SEMI_AUTO. Elle reste volontairement redondante avec
// le veto amont pour qu'une rampe ou un sens memorise dans FB_Translation ne
// puisse alimenter M3 pendant une etape benne.
IF (PRG_03_Modes_Cycle.Data.Auth.Mode = E_Mode.SEMI_AUTO)
   AND NOT M3_CycleTranslationStepAuthorized THEN
    TranslationFinalInterlockRequest.BrakeReleaseRequest := FALSE;
    TranslationFinalInterlockRequest.RequestedDriveControlWord := 0;
    TranslationFinalInterlockRequest.RequestedDriveFreqHz := 0.0;
    TranslationFinalInterlockRequest.ReqTremieSemantic := FALSE;
    TranslationFinalInterlockRequest.ReqMaintenanceSemantic := FALSE;
END_IF;

{endregion}

{region "§4 Publication etat IHM"}
// === 📤 PUBLICATION ÉTAT TRANSLATION IHM (lecture seule) ===
IF instTranslationM3.Fault.Error THEN
    TranslationState.FBState := E_State.ERROR;
ELSIF ABS(instTranslationM3.RequestedDriveFreqHz) > 0.1 THEN
    TranslationState.FBState := E_State.BUSY;
ELSE
    TranslationState.FBState := E_State.READY;
END_IF;
TranslationState.Ready := instTranslationM3.Ready;
TranslationState.Busy := (ABS(instTranslationM3.RequestedDriveFreqHz) > 0.1);
TranslationState.Done := instTranslationM3.TargetReached;
TranslationState.Error := instTranslationM3.Fault.Error;
TranslationState.ErrorId := instTranslationM3.Fault.ErrorId;
TranslationState.BrakeCmd := instTranslationM3.BrakeReleaseRequest;
TranslationState.BrakeCommandOpenConfirmed := instTranslationM3.BrakeCommandOpenConfirmed;
// 🔌 Retour physique direct frein M3 (même source que le SEL §1bis/§2) — consommé FB_TroubleshootingView Idx108
TranslationState.BrakeFeedback := PRG_02_Acquisition.HwIn.Translation.M3_BrakeIsOpen_DI;
TranslationState.PositionReached := instTranslationM3.TargetReached;
TranslationState.DriveControlWord := instTranslationM3.RequestedDriveControlWord;
TranslationState.DriveFreqCmd_Hz := instTranslationM3.RequestedDriveFreqHz;
// 🎯 Cohérence sim : les bits actifs/SpeedCmd_Pct n'affichent la
// consigne QUE si la commande variateur est réellement émise (RequestedDriveControlWord <> 0).
// Sinon, un interlock bloquant (hauteur, SafeStop…) laisserait l'IHM suggérer un mouvement
// qui n'a pas lieu ("je bouge mais ça bouge pas"). Affiche 0 quand c'est bloqué.
TranslationState.ActiveTremie := instTranslationM3.RequestedDriveControlWord = 1;
TranslationState.ActiveMaintenance := instTranslationM3.RequestedDriveControlWord = 2;
TranslationState.SpeedCmd_Pct := SEL(instTranslationM3.RequestedDriveControlWord <> 0, M3_SpeedCmd_Active, 0.0);
TranslationState.PositionTremie := instPosDecoderM3.TranslationPosTremie;
TranslationState.PositionPV := instPosDecoderM3.TranslationPosPV;
TranslationState.PositionP2 := instPosDecoderM3.TranslationPosP2;
TranslationState.PositionP1 := instPosDecoderM3.TranslationPosP1;
TranslationState.PositionMaintenance := instPosDecoderM3.TranslationPosMaintenance;
// Affichage IHM = M3_AtXxxStable (§0quater) — armé sur front
// (direction-dépendant), libéré sur mouvement réel confirmé ≥1.5s (pas juste un rebond capteur
// ni un changement de sens instantané). Même signal que celui consommé par M3_PositionSensorTarget.
TranslationState.AtTremie := M3_AtTremieStable;
TranslationState.AtPV := M3_AtPVStable;
TranslationState.AtP2 := M3_AtP2Stable;
TranslationState.AtP1 := M3_AtP1Stable;
TranslationState.AtMaintenance := M3_AtMaintenanceStable;
// T249-B : "at position" par PLAGE (capteur ON + estime +/-0.5 m) — fiable sans
// dependance frequence variateur, contrairement a AtXxx (front/frequence). + texte statut.
TranslationState.M3StatusText      := M3_StatusText;
TranslationState.EstimatedPosM3_M := instPosEstimatorM3.PositionEstimatedM;
// 📏 T301 — gain odométrique actif + mesure proposée P2 <-> PV (lecture seule, recopie manuelle)
TranslationState.OdometryGainActive := instOdometryGainM3.GainActive;
TranslationState.OdometryCalibValid := instOdometryGainM3.CalibValid;
TranslationState.OdometryMeasureActive := instOdometryGainM3.MeasureActive;
TranslationState.OdometryMeasuredTime_S := instOdometryGainM3.MeasuredTime_S;
TranslationState.OdometryMeasuredFreqAvg_Hz := instOdometryGainM3.MeasuredFreqAvg_Hz;
TranslationState.OdometryMeasuredFreqSpread_Hz := instOdometryGainM3.MeasuredFreqSpread_Hz;
TranslationState.OdometryMeasuredGain := instOdometryGainM3.MeasuredGain;
TranslationState.OdometryMeasureCount := instOdometryGainM3.MeasureCount;
TranslationState.SensorsWord := instPosDecoderM3.SensorsWord;
TranslationState.SensorWordIncoherent := instPosDecoderM3.Incoherent;
TranslationState.LimitSwitchTremie := M3_LimitSwitchTremieStable;
TranslationState.LimitSwitchMaintenance := M3_LimitSwitchMaintenanceStable;
TranslationState.DriveActualFreq_Hz := TO_REAL(PRG_02_Acquisition.Data.M3.ActualFrequencyHz) / 100.0;
TranslationState.DriveThermalOk := PRG_02_Acquisition.HwIn.Translation.M3_ThermalOK_DI;
// 🛡️ Pas de sortie State sur FB_TranslationOutputInterlock : le "vrai état" de la
// barrière finale M3 est dérivé de son défaut (READY normal / ERROR sur défaut barrière).
IF PRG_06_Outputs.instTranslationOutputInterlockM3.Fault.Error THEN
    TranslationState.FinalInterlockState := E_State.ERROR;
ELSE
    TranslationState.FinalInterlockState := E_State.READY;
END_IF;
TranslationState.FinalInterlockReason := PRG_06_Outputs.instTranslationOutputInterlockM3.Reason;
TranslationState.FinalInterlockError := PRG_06_Outputs.instTranslationOutputInterlockM3.Fault.Error;
TranslationState.FinalInterlockErrorId := PRG_06_Outputs.instTranslationOutputInterlockM3.Fault.ErrorId;
TranslationState.FinalBrakeTimeoutElapsed := PRG_06_Outputs.instTranslationOutputInterlockM3.BrakeTimeoutElapsed;
TranslationState.DriveCommReady := (PRG_02_Acquisition.Data.M3.StatusWord AND 16#0080) <> 0;
TranslationState.DrivePowerReady := (PRG_02_Acquisition.Data.M3.StatusWord AND 16#0001) <> 0;
TranslationState.MaintenanceTargetEnable := PRG_03_Modes_Cycle.Data.Auth.MaintenanceM3TargetEnable;
TranslationState.SimulationModeActive := GVL_Simulation.SimulationModeActive;

// 🛡️ Producteur unique (CODE_QUALITY_STANDARDS §5) : la safety M3 (instSafetyTranslationM3)
// est la source de tous les diagnostics de sécurité (ErrorLimitSwitch/ErrorSensorIncoherent).
// Les erreurs propres au mouvement (frein, variateur AC600) restent sur TranslationState.ErrorId
// ci-dessus, bitfield différent, jamais mélangé.
TranslationSafety.SafeStop := M3_SafeStop_Aggregate;
TranslationSafety.PowerCutOff := instSafetyTranslationM3.PowerCutOff;
TranslationSafety.Error := instSafetyTranslationM3.Fault.Error;
TranslationSafety.ErrorId := instSafetyTranslationM3.Fault.ErrorId;
TranslationSafety.LatchedId := instSafetyTranslationM3.Fault.LatchedId;
TranslationSafety.ErrorOperatorComm := instSafetyTranslationM3.ErrorOperatorComm;
TranslationSafety.ErrorDriveComm := instSafetyTranslationM3.ErrorDriveComm;
TranslationSafety.ErrorPhaseRotation := instSafetyTranslationM3.ErrorPhaseRotation;
TranslationSafety.ErrorBrakeThermal := instSafetyTranslationM3.ErrorBrakeThermal;
TranslationSafety.ErrorMecaB := instSafetyTranslationM3.ErrorMecaB;
TranslationSafety.ErrorMecaA := instSafetyTranslationM3.ErrorMecaA;
TranslationSafety.ErrorLimitSwitch := instSafetyTranslationM3.ErrorLimitSwitch;
TranslationSafety.ErrorSensorIncoherent := instSafetyTranslationM3.ErrorSensorIncoherent;
// 🟢 Permis directionnels M3 EFFECTIFS (D1 — Safety AND Process, §1ter) — projetés vers l'IHM
// (source safety : FB_Safety_Translation ; fusion Process en local, modèle treuils PRG_04 §5)
TranslationSafety.EffectivePermitM3_Tremie := EffectivePermitM3_Tremie;
TranslationSafety.EffectivePermitM3_Maintenance := EffectivePermitM3_Maintenance;
TranslationSafety.PowerCutOffSafety := PRG_06_Outputs.M3PowerCutOffSafetyInfo;
TranslationSafety.SafeStopSafety := PRG_06_Outputs.M3SafeStopSafetyInfo;
TranslationSafety.BlockedBySafety := PRG_06_Outputs.M3BlockedBySafetyInfo;

{region "§4bis Trace de blocage terrain M3 (ST_TraceTranslation)"}
// === ↔️ §4bis TRACE DE BLOCAGE TERRAIN M3 (cause priorisée + horodatage) ===
// Diagnostic lecture seule, publié via Data.TranslationTrace et consommé par FB_TroubleshootingView.
// L'ordre IF/ELSIF EST l'ordre de priorité (cf. E_TranslationTraceBlockReason) : la cause la plus
// grave gagne. BlockReasonTimestamp est latched au premier scan du changement (1 scan, mémoire).
// Aucune action de conduite ne dépend de ces champs.
TranslationTrace.SafeStopActive           := M3_SafeStop_Aggregate;
TranslationTrace.SafeStopSourceInput      := M3_SafeStop_Active;
TranslationTrace.SafeStopSourceSafety     := instSafetyTranslationM3.SafeStop;
TranslationTrace.PowerCutOffActive        := instSafetyTranslationM3.PowerCutOff;
TranslationTrace.HeightInterlockBlocking  := NOT M3_HeightInterlockOk;
TranslationTrace.DriveOperational         := PRG_02_Acquisition.Data.Network.DriveM3.Operational;
TranslationTrace.FinalInterlockError      := TranslationState.FinalInterlockError;
// 🟢 Permis directionnels par sens EFFECTIFS (D1 — Safety AND Process, §1ter) — reflet exact des permis appliqués
TranslationTrace.EffectivePermitM3_Tremie      := EffectivePermitM3_Tremie;
TranslationTrace.TremieProcessBlockActive      := M3_TremieProcessBlock;
TranslationTrace.EffectivePermitM3_Maintenance := EffectivePermitM3_Maintenance;

// Permis de mouvement effectif = toutes les barrières levées (agrégat diagnostic)
TranslationTrace.MotionPermitEffective := NOT M3_SafeStop_Aggregate
    AND NOT instSafetyTranslationM3.PowerCutOff
    AND M3_HeightInterlockOk
    AND PRG_02_Acquisition.Data.Network.DriveM3.Operational
    AND NOT TranslationState.FinalInterlockError
    AND NOT instTranslationM3.Fault.Error;

IF instSafetyTranslationM3.PowerCutOff THEN
    TranslationTrace.BlockReason := E_TranslationTraceBlockReason.POWER_CUTOFF;
ELSIF M3_SafeStop_Aggregate THEN
    TranslationTrace.BlockReason := E_TranslationTraceBlockReason.SAFESTOP;
ELSIF instSafetyTranslationM3.Fault.Error THEN
    TranslationTrace.BlockReason := E_TranslationTraceBlockReason.SAFETY_FAULT;
ELSIF NOT M3_HeightInterlockOk THEN
    TranslationTrace.BlockReason := E_TranslationTraceBlockReason.HEIGHT_INTERLOCK;
ELSIF NOT PRG_02_Acquisition.Data.Network.DriveM3.Operational THEN
    TranslationTrace.BlockReason := E_TranslationTraceBlockReason.DRIVE_UNAVAILABLE;
ELSIF TranslationState.FinalInterlockError THEN
    TranslationTrace.BlockReason := E_TranslationTraceBlockReason.FINAL_INTERLOCK;
ELSIF instTranslationM3.Fault.Error THEN
    TranslationTrace.BlockReason := E_TranslationTraceBlockReason.FAULT;
ELSE
    TranslationTrace.BlockReason := E_TranslationTraceBlockReason.NONE;
END_IF;
IF TranslationTrace.BlockReason <> TraceTranslation_PrevReason THEN
    TranslationTrace.BlockReasonTimestamp := TIME_TO_UDINT(TIME());
END_IF;
TraceTranslation_PrevReason := TranslationTrace.BlockReason;
{endregion}

// 🧩 Cause de blocage priorisée sur l'état public IHM (miroir de la trace terrain §4bis)
TranslationState.AxisBlockReason := TranslationTrace.BlockReason;

// === 🔌 PUBLICATION BUS INTER-PRG (Data : ST_TranslationInterPrg) ===
// Copie des structs internes vers le bus de sortie (producteur unique).
Data.TranslationFinalInterlockRequest := TranslationFinalInterlockRequest;
Data.TranslationState                 := TranslationState;
Data.TranslationSafety                := TranslationSafety;
// Arret confirme sur retour reel variateur : la consigne peut deja etre nulle
// pendant la deceleration, elle ne prouve donc pas l'arret physique de M3.
Data.TranslationBusy                  := (ABS(UINT_TO_REAL(PRG_02_Acquisition.Data.M3.ActualFrequencyHz) / 100.0) > 0.5);
Data.TranslationDone                  := instTranslationM3.TargetReached;
Data.M3_AtTremieStable                := M3_AtTremieStable;
Data.M3_AtP1Stable                    := M3_AtP1Stable;
Data.M3_AtMaintenanceStable           := M3_AtMaintenanceStable;
Data.M3_AtWorkPositionStable          := M3_AtWorkPositionStable;
// 🕵️ Trace de blocage terrain (consommée FB_TroubleshootingView)
Data.TranslationTrace                 := TranslationTrace;

{endregion}
END_PROGRAM
